(* IEC 61131-3 sources: volt/packages/volt-lsp-iec/test-corpus/lenze-mid/Device/Plc Logic/Application/Library Manager/L_TT1P_TechnologyModules (part 4) *)

(* ---- L_MB1P_POSPROFILER.pou ---- *)
FUNCTION_BLOCK L_MB1P_POSPROFILER
VAR_INPUT
	XEXECUTE : BOOL;
	XAUXEXECUTE : BOOL;
	XABORT : BOOL;
	XPOSMODE : BOOL;
	ROVERRIDESPEED : REAL;
	ROVERRIDEACC : REAL;
	ROVERRIDEDEC : REAL;
	ROVERRIDEJERKACC : REAL;
	ROVERRIDEJERKDEC : REAL;
	LRACTPOS : LREAL;
	LRACTSPEED : LREAL;
	LRACTACC : LREAL;
	RTASKCYCLE : REAL;
END_VAR
VAR_OUTPUT
	XBUSY : BOOL;
	XDONE : BOOL;
	XABORTED : BOOL;
	XERROR : BOOL;
	LRSETPOS : LREAL;
	LRSETSPEED : LREAL;
	LRSETACC : LREAL;
	DWSTATE : DWORD;
	DWPROFILETYPE : DWORD;
END_VAR
VAR_IN_OUT
	SCPROFILEPARAMETER : L_MB1P_ProfileParameter;
END_VAR
VAR
	SCPROFILEDATA : L_MB1P_ProfileData;
	LREVALTIME : LREAL;
	DWSTATEOFINTERPOLATOR : DWORD;
	XFLAGEXECUTE : BOOL;
	XFLAGAUXEXECUTE : BOOL;
	XFLAGABORT : BOOL;
	SCPROFILEPARAMETERINT : L_MB1P_ProfileParameter;
	ROVERRIDESPEEDOLD : REAL;
	ROVERRIDEACCOLD : REAL;
	ROVERRIDEDECOLD : REAL;
	ROVERRIDEJERKACCOLD : REAL;
	ROVERRIDEJERKDECOLD : REAL;
	XSTARTCALCPROF : BOOL;
	XVELOVEREQZERO : BOOL;
	ARG1 : LREAL;
END_VAR
END_FUNCTION_BLOCK

METHOD CALCPROFILE : BOOL
VAR_INPUT
	DWPROFILETYPE : DWORD;
	LRSTARTACC : LREAL;
	LRSTARTVEL : LREAL;
	SCPROFILEPARAMETER : L_MB1P_ProfileParameter;
	SCMINPROFILEDATA : L_MB1P_IntProfileData;
	SCMAXPROFILEDATA : L_MB1P_IntProfileData;
END_VAR
VAR_OUTPUT
	SCPROFILEDATA : L_MB1P_ProfileData;
	DWSTATE : DWORD;
END_VAR
END_METHOD

METHOD CALCPROFILEDATA : BOOL
VAR_INPUT
	LRSTARTACC : LREAL;
	LRSTARTVEL : LREAL;
	LRSTARTPOS : LREAL;
	XVELMODE : BOOL;
END_VAR
VAR_OUTPUT
	XERROR : BOOL;
	DWSTATE : DWORD;
	DWPROFILETYPE : DWORD;
END_VAR
VAR_IN_OUT
	SCPROFILEDATA : L_MB1P_ProfileData;
	SCPROFILEPARAMETER : L_MB1P_ProfileParameter;
END_VAR
END_METHOD

METHOD IDENTPROFILETYPE : DWORD
VAR_INPUT
	XVELMODE : BOOL;
	LRSTARTACC : LREAL;
	LRSTARTVEL : LREAL;
	SCPROFILEPARAMETER : L_MB1P_ProfileParameter;
END_VAR
VAR_OUTPUT
	DWPROFILETYPE : DWORD;
	SCMINPROFILEDATA : L_MB1P_IntProfileData;
	SCMAXPROFILEDATA : L_MB1P_IntProfileData;
	DWSTATE : DWORD;
END_VAR
END_METHOD

METHOD PROFILEINTERPOLATOR : BOOL
VAR_INPUT
	LREVALTIME : LREAL;
END_VAR
VAR_OUTPUT
	DWSTATE : DWORD;
	LRSETPOS : LREAL;
	LRSETVEL : LREAL;
	LRSETACC : LREAL;
END_VAR
VAR_IN_OUT
	SCPROFILEDATA : L_MB1P_ProfileData;
END_VAR
END_METHOD

METHOD RESETOUTPUT
END_METHOD

METHOD CALCSQRT : LREAL
VAR_INPUT
	ARG1 : LREAL;
END_VAR
END_METHOD

METHOD CALCMINPOSPROFILE : BOOL
VAR_INPUT
	MAXVEL : LREAL;
	MAXACC1 : LREAL;
	MAXACC2 : LREAL;
	JERKACC1 : LREAL;
	JERKACC2 : LREAL;
	RECIPRJERKACC1 : LREAL;
	RECIPRJERKACC2 : LREAL;
	V0_ACC1 : LREAL;
	V0_ACC2 : LREAL;
	A0_ACC1 : LREAL;
	A0_ACC2 : LREAL;
END_VAR
VAR_OUTPUT
	DIMINPOSPROFILETYPE : DINT;
	MINPOSPROFILEDATA : L_MB1P_IntProfileData;
	VMAXMINTRIACC1 : LREAL;
	VMAX_MINTRIACC2 : LREAL;
END_VAR
END_METHOD

METHOD CALCMINPROFILENEGACC : BOOL
VAR_INPUT
	VMAX : LREAL;
	AMAX : LREAL;
	V0 : LREAL;
	A0 : LREAL;
	JERK : LREAL;
	JERKRECIPR : LREAL;
END_VAR
VAR_OUTPUT
	DWPROFILETYPE : DWORD;
	PROFILEDATA_NEGACC : L_MB1P_IntProfileDataAcc;
END_VAR
END_METHOD

METHOD CALCMINPROFILEPOSACC : BOOL
VAR_INPUT
	VMAX : LREAL;
	AMAX : LREAL;
	V0 : LREAL;
	A0 : LREAL;
	JERK : LREAL;
	JERKRECIPR : LREAL;
END_VAR
VAR_OUTPUT
	DWPROFILETYPE : DWORD;
	PROFILEDATA_POSACC : L_MB1P_IntProfileDataAcc;
END_VAR
END_METHOD

METHOD CALCMINTRI : BOOL
VAR_INPUT
	RECIPRJERKACC1 : LREAL;
	RECIPRJERKACC2 : LREAL;
	A0_ACC1 : LREAL;
	V0_ACC1 : LREAL;
	A0_ACC2 : LREAL;
	V0_ACC2 : LREAL;
END_VAR
VAR_OUTPUT
	VMAXMINTRIACC1 : LREAL;
	VMAXMINTRIACC2 : LREAL;
	PROFILEDATA_ACC1 : L_MB1P_IntProfileDataAcc;
	PROFILEDATA_ACC2 : L_MB1P_IntProfileDataAcc;
END_VAR
END_METHOD

METHOD CHECKPROFILEDATA
VAR_INPUT
	DWMODE : DWORD;
	LRTARGETPOS : LREAL;
	LRTARGETVEL : LREAL;
	LRTARGETACC : LREAL;
	LRJERKPHASE7 : LREAL;
END_VAR
VAR_OUTPUT
	XERROR : BOOL;
END_VAR
VAR_IN_OUT
	SCPROFILEDATA : L_MB1P_ProfileData;
END_VAR
END_METHOD

METHOD IDENTMINNEGPROFILE : BOOL
VAR_INPUT
	MINPOSPROFILETYPE : DINT;
	MAXVEL : LREAL;
	MAXACC : LREAL;
	JERK : LREAL;
	RECIPRJERK : LREAL;
	V0_ACC1 : LREAL;
	V0_ACC2 : LREAL;
	A0_ACC1 : LREAL;
	A0_ACC2 : LREAL;
	TARGETPOS : LREAL;
END_VAR
VAR_OUTPUT
	DWPROFILETYPE : DWORD;
END_VAR
VAR_IN_OUT
	SCMAXPROFILEDATA : L_MB1P_IntProfileData;
	SCMINPROFILEDATA : L_MB1P_IntProfileData;
END_VAR
END_METHOD

METHOD IDENTMINPOSPROFILE : BOOL
VAR_INPUT
	MAXVEL : LREAL;
	MAXACC1 : LREAL;
	MAXACC2 : LREAL;
	JERKACC1 : LREAL;
	JERKACC2 : LREAL;
	V0_ACC1 : LREAL;
	V0_ACC2 : LREAL;
	A0_ACC1 : LREAL;
	A0_ACC2 : LREAL;
	TARGETPOS : LREAL;
END_VAR
VAR_OUTPUT
	DWPROFILETYPE : DWORD;
	SCMAXPROFILEDATA : L_MB1P_IntProfileData;
	SCMINPROFILEDATA : L_MB1P_IntProfileData;
END_VAR
END_METHOD

METHOD IDENTSIMPLETRAPNEG : BOOL
VAR_INPUT
	MAXACC2 : LREAL;
	V0_ACC1 : LREAL;
	V0_ACC2 : LREAL;
	A0_ACC1 : LREAL;
	A0_ACC2 : LREAL;
	JERKACC1 : LREAL;
	JERKACC2 : LREAL;
	RECIPRJERKACC2 : LREAL;
	TARGETPOS : LREAL;
END_VAR
VAR_OUTPUT
	DWPROFILETYPE : DWORD;
END_VAR
VAR_IN_OUT
	SCMINPROFILEDATA : L_MB1P_IntProfileData;
	SCMAXPROFILEDATA : L_MB1P_IntProfileData;
END_VAR
END_METHOD

METHOD IDENTSIMPLETRAPPOSTRINEG : BOOL
VAR_INPUT
	MAXACC1 : LREAL;
	JERKACC1 : LREAL;
	RECIPRJERKACC1 : LREAL;
	V0_ACC1 : LREAL;
	A0_ACC1 : LREAL;
	VMAXMINTRIACC1 : LREAL;
	VMAXMINTRIACC2 : LREAL;
	JERKACC2 : LREAL;
	TARGETPOS : LREAL;
END_VAR
VAR_OUTPUT
	DWPROFILETYPE : DWORD;
END_VAR
VAR_IN_OUT
	SCMINPROFILEDATA : L_MB1P_IntProfileData;
	SCMAXPROFILEDATA : L_MB1P_IntProfileData;
END_VAR
END_METHOD

METHOD IDENTSIMPLETRINEG : BOOL
VAR_INPUT
	V0_ACC1 : LREAL;
	A0_ACC1 : LREAL;
	A0_ACC2 : LREAL;
	JERKACC1 : LREAL;
	JERKACC2 : LREAL;
	RECIPRJERKACC2 : LREAL;
	TARGETPOS : LREAL;
END_VAR
VAR_OUTPUT
	DWPROFILETYPE : DWORD;
END_VAR
VAR_IN_OUT
	SCMINPROFILEDATA : L_MB1P_IntProfileData;
	SCMAXPROFILEDATA : L_MB1P_IntProfileData;
END_VAR
END_METHOD

METHOD IDENTSIMPLETRIPOSTRAPNEG : BOOL
VAR_INPUT
	MAXACC2 : LREAL;
	JERKACC2 : LREAL;
	RECIPRJERKACC2 : LREAL;
	V0_ACC2 : LREAL;
	A0_ACC2 : LREAL;
	VMAXMINTRIACC1 : LREAL;
	JERKACC1 : LREAL;
	TARGETPOS : LREAL;
END_VAR
VAR_OUTPUT
	DWPROFILETYPE : DWORD;
END_VAR
VAR_IN_OUT
	SCMINPROFILEDATA : L_MB1P_IntProfileData;
	SCMAXPROFILEDATA : L_MB1P_IntProfileData;
END_VAR
END_METHOD

METHOD IDENTSIMPLETRIPOSTRINEG : BOOL
VAR_INPUT
	V0_ACC1 : LREAL;
	A0_ACC1 : LREAL;
	AMAX : LREAL;
	RECIPRJERKACC1 : LREAL;
	JERKACC1 : LREAL;
	JERKACC2 : LREAL;
	TARGETPOS : LREAL;
	VMAXMINTRIACC1 : LREAL;
	VMAXMINTRIACC2 : LREAL;
END_VAR
VAR_OUTPUT
	DWPROFILETYPE : DWORD;
END_VAR
VAR_IN_OUT
	SCMINPROFILEDATA : L_MB1P_IntProfileData;
	SCMAXPROFILEDATA : L_MB1P_IntProfileData;
END_VAR
END_METHOD

METHOD IDENTTRAPTRI : BOOL
VAR_INPUT
	V_MINTRAPEZACC1 : LREAL;
	MAXACC1 : LREAL;
	JERKACC1 : LREAL;
	JERKACC2 : LREAL;
	A0_ACC1 : LREAL;
	A0_ACC2 : LREAL;
	V0_ACC1 : LREAL;
	V0_ACC2 : LREAL;
	T1_ACC1 : LREAL;
	T3_ACC1 : LREAL;
	DS_1_ACC1 : LREAL;
	TARGETPOS : LREAL;
END_VAR
VAR_OUTPUT
	DWPROFILETYPE : DWORD;
END_VAR
VAR_IN_OUT
	SCMINPROFILEDATA : L_MB1P_IntProfileData;
	SCMAXPROFILEDATA : L_MB1P_IntProfileData;
END_VAR
END_METHOD

METHOD IDENTTRITRAP : BOOL
VAR_INPUT
	V_MINTRAPEZACC2 : LREAL;
	MAXACC2 : LREAL;
	JERKACC1 : LREAL;
	JERKACC2 : LREAL;
	A0_ACC1 : LREAL;
	A0_ACC2 : LREAL;
	V0_ACC1 : LREAL;
	V0_ACC2 : LREAL;
	T1_ACC2 : LREAL;
	T3_ACC2 : LREAL;
	DS_1_ACC2 : LREAL;
	TARGETPOS : LREAL;
END_VAR
VAR_OUTPUT
	DWPROFILETYPE : DWORD;
END_VAR
VAR_IN_OUT
	SCMINPROFILEDATA : L_MB1P_IntProfileData;
	SCMAXPROFILEDATA : L_MB1P_IntProfileData;
END_VAR
END_METHOD

METHOD CALCPROFILE_10A0 : BOOL
VAR_INPUT
	LRSTARTACC : LREAL;
	LRSTARTVEL : LREAL;
	LRMAXACC : LREAL;
	LRMAXDEC : LREAL;
	LRMAXVEL : LREAL;
	LRTARGETACC : LREAL;
	LRTARGETVEL : LREAL;
	LRTARGETPOS : LREAL;
	LRJERKACC : LREAL;
	LRJERKDEC : LREAL;
	LRJERKTIMEACC : LREAL;
	LRJERKTIMEDEC : LREAL;
END_VAR
VAR_OUTPUT
	DWSTATE : DWORD;
END_VAR
VAR_IN_OUT
	SCPROFILEDATA : L_MB1P_ProfileData;
	SCPROFILEPARAMETER : L_MB1P_ProfileParameter;
END_VAR
END_METHOD

METHOD CALCPROFILE_10A0_A0GTAMAX : BOOL
VAR_INPUT
	LRSTARTACC : LREAL;
	LRSTARTVEL : LREAL;
	LRMAXACC : LREAL;
	LRMAXVEL : LREAL;
	LRMAXDEC : LREAL;
	LRTARGETACC : LREAL;
	LRTARGETVEL : LREAL;
	LRTARGETPOS : LREAL;
	LRJERKTIMEACC : LREAL;
	LRJERKTIMEDEC : LREAL;
	LRJERKACC : LREAL;
	LRJERKDEC : LREAL;
END_VAR
VAR_IN_OUT
	SCPROFILEDATA : L_MB1P_ProfileData;
END_VAR
END_METHOD

METHOD CALCPROFILE_10A0_A0LTAMAX : BOOL
VAR_INPUT
	LRSTARTACC : LREAL;
	LRSTARTVEL : LREAL;
	LRMAXACC : LREAL;
	LRMAXVEL : LREAL;
	LRMAXDEC : LREAL;
	LRTARGETACC : LREAL;
	LRTARGETVEL : LREAL;
	LRTARGETPOS : LREAL;
	LRJERKTIMEACC : LREAL;
	LRJERKTIMEDEC : LREAL;
	LRJERKACC : LREAL;
	LRJERKDEC : LREAL;
END_VAR
VAR_IN_OUT
	SCPROFILEDATA : L_MB1P_ProfileData;
END_VAR
END_METHOD

METHOD CALCPROFILE_10B0 : BOOL
VAR_INPUT
	LRSTARTACC : LREAL;
	LRSTARTVEL : LREAL;
	LRMAXACC : LREAL;
	LRMAXDEC : LREAL;
	LRMAXVEL : LREAL;
	LRTARGETACC : LREAL;
	LRTARGETVEL : LREAL;
	LRTARGETPOS : LREAL;
	LRJERKACC : LREAL;
	LRJERKDEC : LREAL;
	LRJERKTIMEACC : LREAL;
	LRJERKTIMEDEC : LREAL;
END_VAR
VAR_OUTPUT
	DWSTATE : DWORD;
END_VAR
VAR_IN_OUT
	SCPROFILEDATA : L_MB1P_ProfileData;
	SCPROFILEPARAMETER : L_MB1P_ProfileParameter;
END_VAR
END_METHOD

METHOD CALCPROFILE_10B0_A0GTAMAX : BOOL
VAR_INPUT
	LRSTARTACC : LREAL;
	LRSTARTVEL : LREAL;
	LRMAXACC : LREAL;
	LRMAXVEL : LREAL;
	LRMAXDEC : LREAL;
	LRTARGETACC : LREAL;
	LRTARGETVEL : LREAL;
	LRTARGETPOS : LREAL;
	LRJERKTIMEACC : LREAL;
	LRJERKTIMEDEC : LREAL;
	LRJERKACC : LREAL;
	LRJERKDEC : LREAL;
END_VAR
VAR_IN_OUT
	SCPROFILEDATA : L_MB1P_ProfileData;
END_VAR
END_METHOD

METHOD CALCPROFILE_10B0_A0LTAMAX : BOOL
VAR_INPUT
	LRSTARTACC : LREAL;
	LRSTARTVEL : LREAL;
	LRMAXACC : LREAL;
	LRMAXVEL : LREAL;
	LRMAXDEC : LREAL;
	LRTARGETACC : LREAL;
	LRTARGETVEL : LREAL;
	LRTARGETPOS : LREAL;
	LRJERKTIMEACC : LREAL;
	LRJERKTIMEDEC : LREAL;
	LRJERKACC : LREAL;
	LRJERKDEC : LREAL;
END_VAR
VAR_IN_OUT
	SCPROFILEDATA : L_MB1P_ProfileData;
END_VAR
END_METHOD

METHOD CALCPROFILE_10C0 : BOOL
VAR_INPUT
	LRSTARTACC : LREAL;
	LRSTARTVEL : LREAL;
	LRMAXACC : LREAL;
	LRMAXDEC : LREAL;
	LRMAXVEL : LREAL;
	LRTARGETACC : LREAL;
	LRTARGETVEL : LREAL;
	LRTARGETPOS : LREAL;
	LRJERKACC : LREAL;
	LRJERKDEC : LREAL;
	LRJERKTIMEACC : LREAL;
	LRJERKTIMEDEC : LREAL;
END_VAR
VAR_OUTPUT
	DWSTATE : DWORD;
END_VAR
VAR_IN_OUT
	SCPROFILEDATA : L_MB1P_ProfileData;
	SCPROFILEPARAMETER : L_MB1P_ProfileParameter;
END_VAR
END_METHOD

METHOD CALCPROFILE_10C0_A0LTAMAXT31 : BOOL
VAR_INPUT
	LRSTARTACC : LREAL;
	LRSTARTVEL : LREAL;
	LRMAXACC : LREAL;
	LRMAXVEL : LREAL;
	LRMAXDEC : LREAL;
	LRTARGETACC : LREAL;
	LRTARGETVEL : LREAL;
	LRTARGETPOS : LREAL;
	LRJERKTIMEACC : LREAL;
	LRJERKTIMEDEC : LREAL;
	LRJERKACC : LREAL;
	LRJERKDEC : LREAL;
END_VAR
VAR_IN_OUT
	SCPROFILEDATA : L_MB1P_ProfileData;
END_VAR
END_METHOD

METHOD CALCPROFILE_10C0_A0LTAMAXT32 : BOOL
VAR_INPUT
	LRSTARTACC : LREAL;
	LRSTARTVEL : LREAL;
	LRMAXACC : LREAL;
	LRMAXVEL : LREAL;
	LRMAXDEC : LREAL;
	LRTARGETACC : LREAL;
	LRTARGETVEL : LREAL;
	LRTARGETPOS : LREAL;
	LRJERKTIMEACC : LREAL;
	LRJERKTIMEDEC : LREAL;
	LRJERKACC : LREAL;
	LRJERKDEC : LREAL;
END_VAR
VAR_IN_OUT
	SCPROFILEDATA : L_MB1P_ProfileData;
END_VAR
END_METHOD

METHOD CALCPROFILE_10D0 : BOOL
VAR_INPUT
	LRSTARTACC : LREAL;
	LRSTARTVEL : LREAL;
	LRMAXACC : LREAL;
	LRMAXDEC : LREAL;
	LRMAXVEL : LREAL;
	LRTARGETACC : LREAL;
	LRTARGETVEL : LREAL;
	LRTARGETPOS : LREAL;
	LRJERKACC : LREAL;
	LRJERKDEC : LREAL;
	LRJERKTIMEACC : LREAL;
	LRJERKTIMEDEC : LREAL;
END_VAR
VAR_OUTPUT
	DWSTATE : DWORD;
END_VAR
VAR_IN_OUT
	SCPROFILEDATA : L_MB1P_ProfileData;
	SCPROFILEPARAMETER : L_MB1P_ProfileParameter;
END_VAR
END_METHOD

METHOD CALCPROFILE_10D0_A0LTAMAXT31T51 : BOOL
VAR_INPUT
	LRSTARTACC : LREAL;
	LRSTARTVEL : LREAL;
	LRMAXACC : LREAL;
	LRMAXVEL : LREAL;
	LRMAXDEC : LREAL;
	LRTARGETACC : LREAL;
	LRTARGETVEL : LREAL;
	LRTARGETPOS : LREAL;
	LRJERKTIMEACC : LREAL;
	LRJERKTIMEDEC : LREAL;
	LRJERKACC : LREAL;
	LRJERKDEC : LREAL;
END_VAR
VAR_IN_OUT
	SCPROFILEDATA : L_MB1P_ProfileData;
END_VAR
END_METHOD

METHOD CALCPROFILE_10D0_A0LTAMAXT31T52 : BOOL
VAR_INPUT
	LRSTARTACC : LREAL;
	LRSTARTVEL : LREAL;
	LRMAXACC : LREAL;
	LRMAXVEL : LREAL;
	LRMAXDEC : LREAL;
	LRTARGETACC : LREAL;
	LRTARGETVEL : LREAL;
	LRTARGETPOS : LREAL;
	LRJERKTIMEACC : LREAL;
	LRJERKTIMEDEC : LREAL;
	LRJERKACC : LREAL;
	LRJERKDEC : LREAL;
END_VAR
VAR_IN_OUT
	SCPROFILEDATA : L_MB1P_ProfileData;
END_VAR
END_METHOD

METHOD CALCPROFILE_10D0_A0LTAMAXT32T51 : BOOL
VAR_INPUT
	LRSTARTACC : LREAL;
	LRSTARTVEL : LREAL;
	LRMAXACC : LREAL;
	LRMAXVEL : LREAL;
	LRMAXDEC : LREAL;
	LRTARGETACC : LREAL;
	LRTARGETVEL : LREAL;
	LRTARGETPOS : LREAL;
	LRJERKTIMEACC : LREAL;
	LRJERKTIMEDEC : LREAL;
	LRJERKACC : LREAL;
	LRJERKDEC : LREAL;
END_VAR
VAR_IN_OUT
	SCPROFILEDATA : L_MB1P_ProfileData;
END_VAR
END_METHOD

METHOD CALCPROFILE_10D0_A0LTAMAXT32T52 : BOOL
VAR_INPUT
	LRSTARTACC : LREAL;
	LRSTARTVEL : LREAL;
	LRMAXACC : LREAL;
	LRMAXVEL : LREAL;
	LRMAXDEC : LREAL;
	LRTARGETACC : LREAL;
	LRTARGETVEL : LREAL;
	LRTARGETPOS : LREAL;
	LRJERKTIMEACC : LREAL;
	LRJERKTIMEDEC : LREAL;
	LRJERKACC : LREAL;
	LRJERKDEC : LREAL;
END_VAR
VAR_IN_OUT
	SCPROFILEDATA : L_MB1P_ProfileData;
END_VAR
END_METHOD

METHOD CALCPROFILE_20A0 : BOOL
VAR_INPUT
	LRSTARTACC : LREAL;
	LRSTARTVEL : LREAL;
	LRMAXACC : LREAL;
	LRMAXDEC : LREAL;
	LRMAXVEL : LREAL;
	LRTARGETACC : LREAL;
	LRTARGETVEL : LREAL;
	LRTARGETPOS : LREAL;
	LRJERKACC : LREAL;
	LRJERKDEC : LREAL;
	LRJERKTIMEACC : LREAL;
	LRJERKTIMEDEC : LREAL;
END_VAR
VAR_OUTPUT
	DWSTATE : DWORD;
END_VAR
VAR_IN_OUT
	SCPROFILEDATA : L_MB1P_ProfileData;
	SCPROFILEPARAMETER : L_MB1P_ProfileParameter;
END_VAR
END_METHOD

METHOD CALCPROFILE_20A0_A0GTAMAXT71 : BOOL
VAR_INPUT
	LRSTARTACC : LREAL;
	LRSTARTVEL : LREAL;
	LRMAXACC : LREAL;
	LRMAXDEC : LREAL;
	LRMAXVEL : LREAL;
	LRTARGETACC : LREAL;
	LRTARGETVEL : LREAL;
	LRTARGETPOS : LREAL;
	LRJERKACC : LREAL;
	LRJERKDEC : LREAL;
	LRJERKTIMEACC : LREAL;
	LRJERKTIMEDEC : LREAL;
END_VAR
VAR_IN_OUT
	SCPROFILEDATA : L_MB1P_ProfileData;
END_VAR
END_METHOD

METHOD CALCPROFILE_20A0_A0GTAMAXT72 : BOOL
VAR_INPUT
	LRSTARTACC : LREAL;
	LRSTARTVEL : LREAL;
	LRMAXACC : LREAL;
	LRMAXDEC : LREAL;
	LRMAXVEL : LREAL;
	LRTARGETACC : LREAL;
	LRTARGETVEL : LREAL;
	LRTARGETPOS : LREAL;
	LRJERKACC : LREAL;
	LRJERKDEC : LREAL;
	LRJERKTIMEACC : LREAL;
	LRJERKTIMEDEC : LREAL;
END_VAR
VAR_IN_OUT
	SCPROFILEDATA : L_MB1P_ProfileData;
END_VAR
END_METHOD

METHOD CALCPROFILE_20A0_A0LTAMAXT71 : BOOL
VAR_INPUT
	LRSTARTACC : LREAL;
	LRSTARTVEL : LREAL;
	LRMAXACC : LREAL;
	LRMAXDEC : LREAL;
	LRMAXVEL : LREAL;
	LRTARGETACC : LREAL;
	LRTARGETVEL : LREAL;
	LRTARGETPOS : LREAL;
	LRJERKACC : LREAL;
	LRJERKDEC : LREAL;
	LRJERKTIMEACC : LREAL;
	LRJERKTIMEDEC : LREAL;
END_VAR
VAR_IN_OUT
	SCPROFILEDATA : L_MB1P_ProfileData;
END_VAR
END_METHOD

METHOD CALCPROFILE_20A0_A0LTAMAXT72 : BOOL
VAR_INPUT
	LRSTARTACC : LREAL;
	LRSTARTVEL : LREAL;
	LRMAXACC : LREAL;
	LRMAXDEC : LREAL;
	LRMAXVEL : LREAL;
	LRTARGETACC : LREAL;
	LRTARGETVEL : LREAL;
	LRTARGETPOS : LREAL;
	LRJERKACC : LREAL;
	LRJERKDEC : LREAL;
	LRJERKTIMEACC : LREAL;
	LRJERKTIMEDEC : LREAL;
END_VAR
VAR_IN_OUT
	SCPROFILEDATA : L_MB1P_ProfileData;
END_VAR
END_METHOD

METHOD CALCPROFILE_20B0 : BOOL
VAR_INPUT
	LRSTARTACC : LREAL;
	LRSTARTVEL : LREAL;
	LRMAXACC : LREAL;
	LRMAXDEC : LREAL;
	LRMAXVEL : LREAL;
	LRTARGETACC : LREAL;
	LRTARGETVEL : LREAL;
	LRTARGETPOS : LREAL;
	LRJERKACC : LREAL;
	LRJERKDEC : LREAL;
	LRJERKTIMEACC : LREAL;
	LRJERKTIMEDEC : LREAL;
	SCMAXPROFILEDATA : L_MB1P_IntProfileData;
	SCMINPROFILEDATA : L_MB1P_IntProfileData;
END_VAR
VAR_OUTPUT
	DWSTATE : DWORD;
END_VAR
VAR_IN_OUT
	SCPROFILEDATA : L_MB1P_ProfileData;
	SCPROFILEPARAMETER : L_MB1P_ProfileParameter;
END_VAR
END_METHOD

METHOD CALCPROFILE_20B0_A0GTAMAXSEARCHTIMEST5T7 : BOOL
VAR_INPUT
	LRSTARTACC : LREAL;
	LRSTARTVEL : LREAL;
	LRMAXACC : LREAL;
	LRMAXDEC : LREAL;
	LRMAXVEL : LREAL;
	LRTARGETACC : LREAL;
	LRTARGETVEL : LREAL;
	LRTARGETPOS : LREAL;
	LRJERKACC : LREAL;
	LRJERKDEC : LREAL;
	LRJERKTIMEACC : LREAL;
	LRJERKTIMEDEC : LREAL;
	T5_STARTVALUE : LREAL;
	T7_STARTVALUE : LREAL;
END_VAR
VAR_OUTPUT
	T5 : LREAL;
	T7 : LREAL;
END_VAR
END_METHOD

METHOD CALCPROFILE_20B0_A0GTAMAXT5T7 : BOOL
VAR_INPUT
	LRSTARTACC : LREAL;
	LRSTARTVEL : LREAL;
	LRMAXACC : LREAL;
	LRMAXDEC : LREAL;
	LRMAXVEL : LREAL;
	LRTARGETACC : LREAL;
	LRTARGETVEL : LREAL;
	LRTARGETPOS : LREAL;
	LRJERKACC : LREAL;
	LRJERKDEC : LREAL;
	LRJERKTIMEACC : LREAL;
	LRJERKTIMEDEC : LREAL;
	T5 : LREAL;
	T7 : LREAL;
END_VAR
VAR_IN_OUT
	SCPROFILEDATA : L_MB1P_ProfileData;
END_VAR
END_METHOD

METHOD CALCPROFILE_20B0_A0LTAMAXSEARCHTIMEST5T7 : BOOL
VAR_INPUT
	LRSTARTACC : LREAL;
	LRSTARTVEL : LREAL;
	LRMAXACC : LREAL;
	LRMAXDEC : LREAL;
	LRMAXVEL : LREAL;
	LRTARGETACC : LREAL;
	LRTARGETVEL : LREAL;
	LRTARGETPOS : LREAL;
	LRJERKACC : LREAL;
	LRJERKDEC : LREAL;
	LRJERKTIMEACC : LREAL;
	LRJERKTIMEDEC : LREAL;
	T5_STARTVALUE : LREAL;
	T7_STARTVALUE : LREAL;
END_VAR
VAR_OUTPUT
	T5 : LREAL;
	T7 : LREAL;
END_VAR
END_METHOD

METHOD CALCPROFILE_20B0_A0LTAMAXT5T7 : BOOL
VAR_INPUT
	LRSTARTACC : LREAL;
	LRSTARTVEL : LREAL;
	LRMAXACC : LREAL;
	LRMAXDEC : LREAL;
	LRMAXVEL : LREAL;
	LRTARGETACC : LREAL;
	LRTARGETVEL : LREAL;
	LRTARGETPOS : LREAL;
	LRJERKACC : LREAL;
	LRJERKDEC : LREAL;
	LRJERKTIMEACC : LREAL;
	LRJERKTIMEDEC : LREAL;
	T5 : LREAL;
	T7 : LREAL;
END_VAR
VAR_IN_OUT
	SCPROFILEDATA : L_MB1P_ProfileData;
END_VAR
END_METHOD

METHOD CALCPROFILE_20BA : BOOL
VAR_INPUT
	LRSTARTACC : LREAL;
	LRSTARTVEL : LREAL;
	LRMAXACC : LREAL;
	LRMAXDEC : LREAL;
	LRMAXVEL : LREAL;
	LRTARGETACC : LREAL;
	LRTARGETVEL : LREAL;
	LRTARGETPOS : LREAL;
	LRJERKACC : LREAL;
	LRJERKDEC : LREAL;
	LRJERKTIMEACC : LREAL;
	LRJERKTIMEDEC : LREAL;
	SCMAXPROFILEDATA : L_MB1P_IntProfileData;
	SCMINPROFILEDATA : L_MB1P_IntProfileData;
END_VAR
VAR_OUTPUT
	DWSTATE : DWORD;
END_VAR
VAR_IN_OUT
	SCPROFILEDATA : L_MB1P_ProfileData;
	SCPROFILEPARAMETER : L_MB1P_ProfileParameter;
END_VAR
END_METHOD

METHOD CALCPROFILE_20BA_A0GTAMAX : BOOL
VAR_INPUT
	LRSTARTACC : LREAL;
	LRSTARTVEL : LREAL;
	LRMAXACC : LREAL;
	LRMAXDEC : LREAL;
	LRMAXVEL : LREAL;
	LRTARGETACC : LREAL;
	LRTARGETVEL : LREAL;
	LRTARGETPOS : LREAL;
	LRJERKACC : LREAL;
	LRJERKDEC : LREAL;
	LRJERKTIMEACC : LREAL;
	LRJERKTIMEDEC : LREAL;
	T7 : LREAL;
END_VAR
VAR_IN_OUT
	SCPROFILEDATA : L_MB1P_ProfileData;
END_VAR
END_METHOD

METHOD CALCPROFILE_20BA_A0LETAMAX : BOOL
VAR_INPUT
	LRSTARTACC : LREAL;
	LRSTARTVEL : LREAL;
	LRMAXACC : LREAL;
	LRMAXDEC : LREAL;
	LRMAXVEL : LREAL;
	LRTARGETACC : LREAL;
	LRTARGETVEL : LREAL;
	LRTARGETPOS : LREAL;
	LRJERKACC : LREAL;
	LRJERKDEC : LREAL;
	LRJERKTIMEACC : LREAL;
	LRJERKTIMEDEC : LREAL;
	T7 : LREAL;
END_VAR
VAR_IN_OUT
	SCPROFILEDATA : L_MB1P_ProfileData;
END_VAR
END_METHOD

METHOD CALCPROFILE_20BA_AOGTAMAX_SEARCHTIMES : BOOL
VAR_INPUT
	LRSTARTACC : LREAL;
	LRSTARTVEL : LREAL;
	LRMAXACC : LREAL;
	LRMAXDEC : LREAL;
	LRMAXVEL : LREAL;
	LRTARGETACC : LREAL;
	LRTARGETVEL : LREAL;
	LRTARGETPOS : LREAL;
	LRJERKACC : LREAL;
	LRJERKDEC : LREAL;
	LRJERKTIMEACC : LREAL;
	LRJERKTIMEDEC : LREAL;
	T7_MINVALUE : LREAL;
	T7_MAXVALUE : LREAL;
END_VAR
VAR_OUTPUT
	T7 : LREAL;
END_VAR
END_METHOD

METHOD CALCPROFILE_20BA_AOLETAMAX_SEARCHTIMES : BOOL
VAR_INPUT
	LRSTARTACC : LREAL;
	LRSTARTVEL : LREAL;
	LRMAXACC : LREAL;
	LRMAXDEC : LREAL;
	LRMAXVEL : LREAL;
	LRTARGETACC : LREAL;
	LRTARGETVEL : LREAL;
	LRTARGETPOS : LREAL;
	LRJERKACC : LREAL;
	LRJERKDEC : LREAL;
	LRJERKTIMEACC : LREAL;
	LRJERKTIMEDEC : LREAL;
	T7_MINVALUE : LREAL;
	T7_MAXVALUE : LREAL;
END_VAR
VAR_OUTPUT
	T7 : LREAL;
END_VAR
END_METHOD

METHOD CALCPROFILE_20C0 : BOOL
VAR_INPUT
	LRSTARTACC : LREAL;
	LRSTARTVEL : LREAL;
	LRMAXACC : LREAL;
	LRMAXDEC : LREAL;
	LRMAXVEL : LREAL;
	LRTARGETACC : LREAL;
	LRTARGETVEL : LREAL;
	LRTARGETPOS : LREAL;
	LRJERKACC : LREAL;
	LRJERKDEC : LREAL;
	LRJERKTIMEACC : LREAL;
	LRJERKTIMEDEC : LREAL;
	SCMAXPROFILEDATA : L_MB1P_IntProfileData;
	SCMINPROFILEDATA : L_MB1P_IntProfileData;
END_VAR
VAR_OUTPUT
	DWSTATE : DWORD;
END_VAR
VAR_IN_OUT
	SCPROFILEDATA : L_MB1P_ProfileData;
	SCPROFILEPARAMETER : L_MB1P_ProfileParameter;
END_VAR
END_METHOD

METHOD CALCPROFILE_20C0_SEARCHTIMEST5T7 : BOOL
VAR_INPUT
	LRSTARTACC : LREAL;
	LRSTARTVEL : LREAL;
	LRMAXACC : LREAL;
	LRMAXDEC : LREAL;
	LRMAXVEL : LREAL;
	LRTARGETACC : LREAL;
	LRTARGETVEL : LREAL;
	LRTARGETPOS : LREAL;
	LRJERKACC : LREAL;
	LRJERKDEC : LREAL;
	LRJERKTIMEACC : LREAL;
	LRJERKTIMEDEC : LREAL;
	T5_STARTVALUE : LREAL;
	T7_STARTVALUE : LREAL;
END_VAR
VAR_OUTPUT
	T5 : LREAL;
	T7 : LREAL;
END_VAR
END_METHOD

METHOD CALCPROFILE_20C0_AELTAMAXT5T7 : BOOL
VAR_INPUT
	LRSTARTACC : LREAL;
	LRSTARTVEL : LREAL;
	LRMAXACC : LREAL;
	LRMAXDEC : LREAL;
	LRMAXVEL : LREAL;
	LRTARGETACC : LREAL;
	LRTARGETVEL : LREAL;
	LRTARGETPOS : LREAL;
	LRJERKACC : LREAL;
	LRJERKDEC : LREAL;
	LRJERKTIMEACC : LREAL;
	LRJERKTIMEDEC : LREAL;
	T5 : LREAL;
	T7 : LREAL;
END_VAR
VAR_IN_OUT
	SCPROFILEDATA : L_MB1P_ProfileData;
END_VAR
END_METHOD

METHOD CALCPROFILE_20CB : BOOL
VAR_INPUT
	LRSTARTACC : LREAL;
	LRSTARTVEL : LREAL;
	LRMAXACC : LREAL;
	LRMAXDEC : LREAL;
	LRMAXVEL : LREAL;
	LRTARGETACC : LREAL;
	LRTARGETVEL : LREAL;
	LRTARGETPOS : LREAL;
	LRJERKACC : LREAL;
	LRJERKDEC : LREAL;
	LRJERKTIMEACC : LREAL;
	LRJERKTIMEDEC : LREAL;
	SCMAXPROFILEDATA : L_MB1P_IntProfileData;
	SCMINPROFILEDATA : L_MB1P_IntProfileData;
END_VAR
VAR_OUTPUT
	DWSTATE : DWORD;
END_VAR
VAR_IN_OUT
	SCPROFILEDATA : L_MB1P_ProfileData;
	SCPROFILEPARAMETER : L_MB1P_ProfileParameter;
END_VAR
END_METHOD

METHOD CALCPROFILE_20CB_AOGET0 : BOOL
VAR_INPUT
	LRSTARTACC : LREAL;
	LRSTARTVEL : LREAL;
	LRMAXACC : LREAL;
	LRMAXDEC : LREAL;
	LRMAXVEL : LREAL;
	LRTARGETACC : LREAL;
	LRTARGETVEL : LREAL;
	LRTARGETPOS : LREAL;
	LRJERKACC : LREAL;
	LRJERKDEC : LREAL;
	LRJERKTIMEACC : LREAL;
	LRJERKTIMEDEC : LREAL;
	T7 : LREAL;
END_VAR
VAR_IN_OUT
	SCPROFILEDATA : L_MB1P_ProfileData;
END_VAR
END_METHOD

METHOD CALCPROFILE_20CB_AOLT0 : BOOL
VAR_INPUT
	LRSTARTACC : LREAL;
	LRSTARTVEL : LREAL;
	LRMAXACC : LREAL;
	LRMAXDEC : LREAL;
	LRMAXVEL : LREAL;
	LRTARGETACC : LREAL;
	LRTARGETVEL : LREAL;
	LRTARGETPOS : LREAL;
	LRJERKACC : LREAL;
	LRJERKDEC : LREAL;
	LRJERKTIMEACC : LREAL;
	LRJERKTIMEDEC : LREAL;
	T7 : LREAL;
END_VAR
VAR_IN_OUT
	SCPROFILEDATA : L_MB1P_ProfileData;
END_VAR
END_METHOD

METHOD CALCPROFILE_20CBAOGET0_SEARCHTIMES : BOOL
VAR_INPUT
	LRSTARTACC : LREAL;
	LRSTARTVEL : LREAL;
	LRMAXACC : LREAL;
	LRMAXDEC : LREAL;
	LRMAXVEL : LREAL;
	LRTARGETACC : LREAL;
	LRTARGETVEL : LREAL;
	LRTARGETPOS : LREAL;
	LRJERKACC : LREAL;
	LRJERKDEC : LREAL;
	LRJERKTIMEACC : LREAL;
	LRJERKTIMEDEC : LREAL;
	T7_MINVALUE : LREAL;
	T7_MAXVALUE : LREAL;
END_VAR
VAR_OUTPUT
	T7 : LREAL;
END_VAR
END_METHOD

METHOD CALCPROFILE_20CBAOLT0_SEARCHTIMES : BOOL
VAR_INPUT
	LRSTARTACC : LREAL;
	LRSTARTVEL : LREAL;
	LRMAXACC : LREAL;
	LRMAXDEC : LREAL;
	LRMAXVEL : LREAL;
	LRTARGETACC : LREAL;
	LRTARGETVEL : LREAL;
	LRTARGETPOS : LREAL;
	LRJERKACC : LREAL;
	LRJERKDEC : LREAL;
	LRJERKTIMEACC : LREAL;
	LRJERKTIMEDEC : LREAL;
	T7_MINVALUE : LREAL;
	T7_MAXVALUE : LREAL;
END_VAR
VAR_OUTPUT
	T7 : LREAL;
END_VAR
END_METHOD

METHOD CALCPROFILE_20D0 : BOOL
VAR_INPUT
	LRSTARTACC : LREAL;
	LRSTARTVEL : LREAL;
	LRMAXACC : LREAL;
	LRMAXDEC : LREAL;
	LRMAXVEL : LREAL;
	LRTARGETACC : LREAL;
	LRTARGETVEL : LREAL;
	LRTARGETPOS : LREAL;
	LRJERKACC : LREAL;
	LRJERKDEC : LREAL;
	LRJERKTIMEACC : LREAL;
	LRJERKTIMEDEC : LREAL;
	SCMAXPROFILEDATA : L_MB1P_IntProfileData;
	SCMINPROFILEDATA : L_MB1P_IntProfileData;
END_VAR
VAR_OUTPUT
	DWSTATE : DWORD;
END_VAR
VAR_IN_OUT
	SCPROFILEDATA : L_MB1P_ProfileData;
	SCPROFILEPARAMETER : L_MB1P_ProfileParameter;
END_VAR
END_METHOD

METHOD CALCPROFILE_20D0_SEARCHTIMEST5T7 : BOOL
VAR_INPUT
	LRSTARTACC : LREAL;
	LRSTARTVEL : LREAL;
	LRMAXACC : LREAL;
	LRMAXDEC : LREAL;
	LRMAXVEL : LREAL;
	LRTARGETACC : LREAL;
	LRTARGETVEL : LREAL;
	LRTARGETPOS : LREAL;
	LRJERKACC : LREAL;
	LRJERKDEC : LREAL;
	LRJERKTIMEACC : LREAL;
	LRJERKTIMEDEC : LREAL;
	T5_STARTVALUE : LREAL;
	T7_STARTVALUE : LREAL;
END_VAR
VAR_OUTPUT
	T5 : LREAL;
	T7 : LREAL;
END_VAR
END_METHOD

METHOD CALCPROFILE_20D0_A0LTAMAXT5T7 : BOOL
VAR_INPUT
	LRSTARTACC : LREAL;
	LRSTARTVEL : LREAL;
	LRMAXACC : LREAL;
	LRMAXDEC : LREAL;
	LRMAXVEL : LREAL;
	LRTARGETACC : LREAL;
	LRTARGETVEL : LREAL;
	LRTARGETPOS : LREAL;
	LRJERKACC : LREAL;
	LRJERKDEC : LREAL;
	LRJERKTIMEACC : LREAL;
	LRJERKTIMEDEC : LREAL;
	T5 : LREAL;
	T7 : LREAL;
END_VAR
VAR_IN_OUT
	SCPROFILEDATA : L_MB1P_ProfileData;
END_VAR
END_METHOD

METHOD CALCPROFILE_20D1 : BOOL
VAR_INPUT
	LRSTARTACC : LREAL;
	LRSTARTVEL : LREAL;
	LRMAXACC : LREAL;
	LRMAXDEC : LREAL;
	LRMAXVEL : LREAL;
	LRTARGETACC : LREAL;
	LRTARGETVEL : LREAL;
	LRTARGETPOS : LREAL;
	LRJERKACC : LREAL;
	LRJERKDEC : LREAL;
	LRJERKTIMEACC : LREAL;
	LRJERKTIMEDEC : LREAL;
	SCMAXPROFILEDATA : L_MB1P_IntProfileData;
	SCMINPROFILEDATA : L_MB1P_IntProfileData;
END_VAR
VAR_OUTPUT
	DWSTATE : DWORD;
END_VAR
VAR_IN_OUT
	SCPROFILEDATA : L_MB1P_ProfileData;
	SCPROFILEPARAMETER : L_MB1P_ProfileParameter;
END_VAR
END_METHOD

METHOD CALCPROFILE_20D1_AOGET0 : BOOL
VAR_INPUT
	LRSTARTACC : LREAL;
	LRSTARTVEL : LREAL;
	LRMAXACC : LREAL;
	LRMAXDEC : LREAL;
	LRMAXVEL : LREAL;
	LRTARGETACC : LREAL;
	LRTARGETVEL : LREAL;
	LRTARGETPOS : LREAL;
	LRJERKACC : LREAL;
	LRJERKDEC : LREAL;
	LRJERKTIMEACC : LREAL;
	LRJERKTIMEDEC : LREAL;
	T7 : LREAL;
END_VAR
VAR_IN_OUT
	SCPROFILEDATA : L_MB1P_ProfileData;
END_VAR
END_METHOD

METHOD CALCPROFILE_20D1_AOLT0 : BOOL
VAR_INPUT
	LRSTARTACC : LREAL;
	LRSTARTVEL : LREAL;
	LRMAXACC : LREAL;
	LRMAXDEC : LREAL;
	LRMAXVEL : LREAL;
	LRTARGETACC : LREAL;
	LRTARGETVEL : LREAL;
	LRTARGETPOS : LREAL;
	LRJERKACC : LREAL;
	LRJERKDEC : LREAL;
	LRJERKTIMEACC : LREAL;
	LRJERKTIMEDEC : LREAL;
	T7 : LREAL;
END_VAR
VAR_IN_OUT
	SCPROFILEDATA : L_MB1P_ProfileData;
END_VAR
END_METHOD

METHOD CALCPROFILE_20D1AOGET0_SEARCHTIMES : BOOL
VAR_INPUT
	LRSTARTACC : LREAL;
	LRSTARTVEL : LREAL;
	LRMAXACC : LREAL;
	LRMAXDEC : LREAL;
	LRMAXVEL : LREAL;
	LRTARGETACC : LREAL;
	LRTARGETVEL : LREAL;
	LRTARGETPOS : LREAL;
	LRJERKACC : LREAL;
	LRJERKDEC : LREAL;
	LRJERKTIMEACC : LREAL;
	LRJERKTIMEDEC : LREAL;
	T7_STARTVALUE : LREAL;
END_VAR
VAR_OUTPUT
	T7 : LREAL;
END_VAR
END_METHOD

METHOD CALCPROFILE_20D1AOLT0_SEARCHTIMES : BOOL
VAR_INPUT
	LRSTARTACC : LREAL;
	LRSTARTVEL : LREAL;
	LRMAXACC : LREAL;
	LRMAXDEC : LREAL;
	LRMAXVEL : LREAL;
	LRTARGETACC : LREAL;
	LRTARGETVEL : LREAL;
	LRTARGETPOS : LREAL;
	LRJERKACC : LREAL;
	LRJERKDEC : LREAL;
	LRJERKTIMEACC : LREAL;
	LRJERKTIMEDEC : LREAL;
	T7_STARTVALUE : LREAL;
END_VAR
VAR_OUTPUT
	T7 : LREAL;
END_VAR
END_METHOD

METHOD CALCPROFILE_20DA : BOOL
VAR_INPUT
	LRSTARTACC : LREAL;
	LRSTARTVEL : LREAL;
	LRMAXACC : LREAL;
	LRMAXDEC : LREAL;
	LRMAXVEL : LREAL;
	LRTARGETACC : LREAL;
	LRTARGETVEL : LREAL;
	LRTARGETPOS : LREAL;
	LRJERKACC : LREAL;
	LRJERKDEC : LREAL;
	LRJERKTIMEACC : LREAL;
	LRJERKTIMEDEC : LREAL;
	SCMAXPROFILEDATA : L_MB1P_IntProfileData;
	SCMINPROFILEDATA : L_MB1P_IntProfileData;
END_VAR
VAR_OUTPUT
	DWSTATE : DWORD;
END_VAR
VAR_IN_OUT
	SCPROFILEDATA : L_MB1P_ProfileData;
	SCPROFILEPARAMETER : L_MB1P_ProfileParameter;
END_VAR
END_METHOD

METHOD CALCPROFILE_20DA_AELT0 : BOOL
VAR_INPUT
	LRSTARTACC : LREAL;
	LRSTARTVEL : LREAL;
	LRMAXACC : LREAL;
	LRMAXDEC : LREAL;
	LRMAXVEL : LREAL;
	LRTARGETACC : LREAL;
	LRTARGETVEL : LREAL;
	LRTARGETPOS : LREAL;
	LRJERKACC : LREAL;
	LRJERKDEC : LREAL;
	LRJERKTIMEACC : LREAL;
	LRJERKTIMEDEC : LREAL;
	T7 : LREAL;
END_VAR
VAR_IN_OUT
	SCPROFILEDATA : L_MB1P_ProfileData;
END_VAR
END_METHOD

METHOD CALCPROFILE_20DAAELT0_SEARCHTIMES : BOOL
VAR_INPUT
	LRSTARTACC : LREAL;
	LRSTARTVEL : LREAL;
	LRMAXACC : LREAL;
	LRMAXDEC : LREAL;
	LRMAXVEL : LREAL;
	LRTARGETACC : LREAL;
	LRTARGETVEL : LREAL;
	LRTARGETPOS : LREAL;
	LRJERKACC : LREAL;
	LRJERKDEC : LREAL;
	LRJERKTIMEACC : LREAL;
	LRJERKTIMEDEC : LREAL;
	T7_MINVALUE : LREAL;
	T7_MAXVALUE : LREAL;
END_VAR
VAR_OUTPUT
	T7 : LREAL;
END_VAR
END_METHOD

METHOD CALCPROFILE_20DB : BOOL
VAR_INPUT
	LRSTARTACC : LREAL;
	LRSTARTVEL : LREAL;
	LRMAXACC : LREAL;
	LRMAXDEC : LREAL;
	LRMAXVEL : LREAL;
	LRTARGETACC : LREAL;
	LRTARGETVEL : LREAL;
	LRTARGETPOS : LREAL;
	LRJERKACC : LREAL;
	LRJERKDEC : LREAL;
	LRJERKTIMEACC : LREAL;
	LRJERKTIMEDEC : LREAL;
	SCMAXPROFILEDATA : L_MB1P_IntProfileData;
	SCMINPROFILEDATA : L_MB1P_IntProfileData;
END_VAR
VAR_OUTPUT
	DWSTATE : DWORD;
END_VAR
VAR_IN_OUT
	SCPROFILEDATA : L_MB1P_ProfileData;
	SCPROFILEPARAMETER : L_MB1P_ProfileParameter;
END_VAR
END_METHOD

METHOD CALCPROFILE_20DB_AOGET0 : BOOL
VAR_INPUT
	LRSTARTACC : LREAL;
	LRSTARTVEL : LREAL;
	LRMAXACC : LREAL;
	LRMAXDEC : LREAL;
	LRMAXVEL : LREAL;
	LRTARGETACC : LREAL;
	LRTARGETVEL : LREAL;
	LRTARGETPOS : LREAL;
	LRJERKACC : LREAL;
	LRJERKDEC : LREAL;
	LRJERKTIMEACC : LREAL;
	LRJERKTIMEDEC : LREAL;
	T7 : LREAL;
END_VAR
VAR_IN_OUT
	SCPROFILEDATA : L_MB1P_ProfileData;
END_VAR
END_METHOD

METHOD CALCPROFILE_20DB_AOLT0 : BOOL
VAR_INPUT
	LRSTARTACC : LREAL;
	LRSTARTVEL : LREAL;
	LRMAXACC : LREAL;
	LRMAXDEC : LREAL;
	LRMAXVEL : LREAL;
	LRTARGETACC : LREAL;
	LRTARGETVEL : LREAL;
	LRTARGETPOS : LREAL;
	LRJERKACC : LREAL;
	LRJERKDEC : LREAL;
	LRJERKTIMEACC : LREAL;
	LRJERKTIMEDEC : LREAL;
	T7 : LREAL;
END_VAR
VAR_IN_OUT
	SCPROFILEDATA : L_MB1P_ProfileData;
END_VAR
END_METHOD

METHOD CALCPROFILE_20DBAOGET0_SEARCHTIMES : BOOL
VAR_INPUT
	LRSTARTACC : LREAL;
	LRSTARTVEL : LREAL;
	LRMAXACC : LREAL;
	LRMAXDEC : LREAL;
	LRMAXVEL : LREAL;
	LRTARGETACC : LREAL;
	LRTARGETVEL : LREAL;
	LRTARGETPOS : LREAL;
	LRJERKACC : LREAL;
	LRJERKDEC : LREAL;
	LRJERKTIMEACC : LREAL;
	LRJERKTIMEDEC : LREAL;
	T7_MINVALUE : LREAL;
	T7_MAXVALUE : LREAL;
END_VAR
VAR_OUTPUT
	T7 : LREAL;
END_VAR
END_METHOD

METHOD CALCPROFILE_20DBAOLT0_SEARCHTIMES : BOOL
VAR_INPUT
	LRSTARTACC : LREAL;
	LRSTARTVEL : LREAL;
	LRMAXACC : LREAL;
	LRMAXDEC : LREAL;
	LRMAXVEL : LREAL;
	LRTARGETACC : LREAL;
	LRTARGETVEL : LREAL;
	LRTARGETPOS : LREAL;
	LRJERKACC : LREAL;
	LRJERKDEC : LREAL;
	LRJERKTIMEACC : LREAL;
	LRJERKTIMEDEC : LREAL;
	T7_MINVALUE : LREAL;
	T7_MAXVALUE : LREAL;
END_VAR
VAR_OUTPUT
	T7 : LREAL;
END_VAR
END_METHOD

METHOD CALCPROFILE_30A0 : BOOL
VAR_INPUT
	LRSTARTACC : LREAL;
	LRSTARTVEL : LREAL;
	LRMAXACC : LREAL;
	LRMAXDEC : LREAL;
	LRMAXVEL : LREAL;
	LRTARGETACC : LREAL;
	LRTARGETVEL : LREAL;
	LRTARGETPOS : LREAL;
	LRJERKACC : LREAL;
	LRJERKDEC : LREAL;
	LRJERKTIMEACC : LREAL;
	LRJERKTIMEDEC : LREAL;
END_VAR
VAR_OUTPUT
	DWSTATE : DWORD;
END_VAR
VAR_IN_OUT
	SCPROFILEDATA : L_MB1P_ProfileData;
	SCPROFILEPARAMETER : L_MB1P_ProfileParameter;
END_VAR
END_METHOD

METHOD CALCPROFILE_30A0_A0GTAMAX : BOOL
VAR_INPUT
	LRSTARTACC : LREAL;
	LRSTARTVEL : LREAL;
	LRMAXACC : LREAL;
	LRMAXDEC : LREAL;
	LRMAXVEL : LREAL;
	LRTARGETACC : LREAL;
	LRTARGETVEL : LREAL;
	LRTARGETPOS : LREAL;
	LRJERKACC : LREAL;
	LRJERKDEC : LREAL;
	LRJERKTIMEACC : LREAL;
	LRJERKTIMEDEC : LREAL;
END_VAR
VAR_IN_OUT
	SCPROFILEDATA : L_MB1P_ProfileData;
END_VAR
END_METHOD

METHOD CALCPROFILE_30A0_A0LTAMAX : BOOL
VAR_INPUT
	LRSTARTACC : LREAL;
	LRSTARTVEL : LREAL;
	LRMAXACC : LREAL;
	LRMAXDEC : LREAL;
	LRMAXVEL : LREAL;
	LRTARGETACC : LREAL;
	LRTARGETVEL : LREAL;
	LRTARGETPOS : LREAL;
	LRJERKACC : LREAL;
	LRJERKDEC : LREAL;
	LRJERKTIMEACC : LREAL;
	LRJERKTIMEDEC : LREAL;
END_VAR
VAR_IN_OUT
	SCPROFILEDATA : L_MB1P_ProfileData;
END_VAR
END_METHOD

METHOD CALCPROFILE_30B0 : BOOL
VAR_INPUT
	LRSTARTACC : LREAL;
	LRSTARTVEL : LREAL;
	LRMAXACC : LREAL;
	LRMAXDEC : LREAL;
	LRMAXVEL : LREAL;
	LRTARGETACC : LREAL;
	LRTARGETVEL : LREAL;
	LRTARGETPOS : LREAL;
	LRJERKACC : LREAL;
	LRJERKDEC : LREAL;
	LRJERKTIMEACC : LREAL;
	LRJERKTIMEDEC : LREAL;
END_VAR
VAR_OUTPUT
	DWSTATE : DWORD;
END_VAR
VAR_IN_OUT
	SCPROFILEDATA : L_MB1P_ProfileData;
	SCPROFILEPARAMETER : L_MB1P_ProfileParameter;
END_VAR
END_METHOD

METHOD CALCPROFILE_30B0_A0GTAMAXT51 : BOOL
VAR_INPUT
	LRSTARTACC : LREAL;
	LRSTARTVEL : LREAL;
	LRMAXACC : LREAL;
	LRMAXDEC : LREAL;
	LRMAXVEL : LREAL;
	LRTARGETACC : LREAL;
	LRTARGETVEL : LREAL;
	LRTARGETPOS : LREAL;
	LRJERKACC : LREAL;
	LRJERKDEC : LREAL;
	LRJERKTIMEACC : LREAL;
	LRJERKTIMEDEC : LREAL;
END_VAR
VAR_IN_OUT
	SCPROFILEDATA : L_MB1P_ProfileData;
END_VAR
END_METHOD

METHOD CALCPROFILE_30B0_A0GTAMAXT52 : BOOL
VAR_INPUT
	LRSTARTACC : LREAL;
	LRSTARTVEL : LREAL;
	LRMAXACC : LREAL;
	LRMAXDEC : LREAL;
	LRMAXVEL : LREAL;
	LRTARGETACC : LREAL;
	LRTARGETVEL : LREAL;
	LRTARGETPOS : LREAL;
	LRJERKACC : LREAL;
	LRJERKDEC : LREAL;
	LRJERKTIMEACC : LREAL;
	LRJERKTIMEDEC : LREAL;
END_VAR
VAR_IN_OUT
	SCPROFILEDATA : L_MB1P_ProfileData;
END_VAR
END_METHOD

METHOD CALCPROFILE_30B0_A0LTAMAXT51 : BOOL
VAR_INPUT
	LRSTARTACC : LREAL;
	LRSTARTVEL : LREAL;
	LRMAXACC : LREAL;
	LRMAXDEC : LREAL;
	LRMAXVEL : LREAL;
	LRTARGETACC : LREAL;
	LRTARGETVEL : LREAL;
	LRTARGETPOS : LREAL;
	LRJERKACC : LREAL;
	LRJERKDEC : LREAL;
	LRJERKTIMEACC : LREAL;
	LRJERKTIMEDEC : LREAL;
END_VAR
VAR_IN_OUT
	SCPROFILEDATA : L_MB1P_ProfileData;
END_VAR
END_METHOD

METHOD CALCPROFILE_30B0_A0LTAMAXT52 : BOOL
VAR_INPUT
	LRSTARTACC : LREAL;
	LRSTARTVEL : LREAL;
	LRMAXACC : LREAL;
	LRMAXDEC : LREAL;
	LRMAXVEL : LREAL;
	LRTARGETACC : LREAL;
	LRTARGETVEL : LREAL;
	LRTARGETPOS : LREAL;
	LRJERKACC : LREAL;
	LRJERKDEC : LREAL;
	LRJERKTIMEACC : LREAL;
	LRJERKTIMEDEC : LREAL;
END_VAR
VAR_IN_OUT
	SCPROFILEDATA : L_MB1P_ProfileData;
END_VAR
END_METHOD

METHOD CALCPROFILE_30C0 : BOOL
VAR_INPUT
	LRSTARTACC : LREAL;
	LRSTARTVEL : LREAL;
	LRMAXACC : LREAL;
	LRMAXDEC : LREAL;
	LRMAXVEL : LREAL;
	LRTARGETACC : LREAL;
	LRTARGETVEL : LREAL;
	LRTARGETPOS : LREAL;
	LRJERKACC : LREAL;
	LRJERKDEC : LREAL;
	LRJERKTIMEACC : LREAL;
	LRJERKTIMEDEC : LREAL;
END_VAR
VAR_OUTPUT
	DWSTATE : DWORD;
END_VAR
VAR_IN_OUT
	SCPROFILEDATA : L_MB1P_ProfileData;
	SCPROFILEPARAMETER : L_MB1P_ProfileParameter;
END_VAR
END_METHOD

METHOD CALCPROFILE_30C0_A0GTAMAXT31 : BOOL
VAR_INPUT
	LRSTARTACC : LREAL;
	LRSTARTVEL : LREAL;
	LRMAXACC : LREAL;
	LRMAXDEC : LREAL;
	LRMAXVEL : LREAL;
	LRTARGETACC : LREAL;
	LRTARGETVEL : LREAL;
	LRTARGETPOS : LREAL;
	LRJERKACC : LREAL;
	LRJERKDEC : LREAL;
	LRJERKTIMEACC : LREAL;
	LRJERKTIMEDEC : LREAL;
END_VAR
VAR_IN_OUT
	SCPROFILEDATA : L_MB1P_ProfileData;
END_VAR
END_METHOD

METHOD CALCPROFILE_30C0_A0GTAMAXT32 : BOOL
VAR_INPUT
	LRSTARTACC : LREAL;
	LRSTARTVEL : LREAL;
	LRMAXACC : LREAL;
	LRMAXDEC : LREAL;
	LRMAXVEL : LREAL;
	LRTARGETACC : LREAL;
	LRTARGETVEL : LREAL;
	LRTARGETPOS : LREAL;
	LRJERKACC : LREAL;
	LRJERKDEC : LREAL;
	LRJERKTIMEACC : LREAL;
	LRJERKTIMEDEC : LREAL;
END_VAR
VAR_IN_OUT
	SCPROFILEDATA : L_MB1P_ProfileData;
END_VAR
END_METHOD

METHOD CALCPROFILE_30CB : BOOL
VAR_INPUT
	LRSTARTACC : LREAL;
	LRSTARTVEL : LREAL;
	LRMAXACC : LREAL;
	LRMAXDEC : LREAL;
	LRMAXVEL : LREAL;
	LRTARGETACC : LREAL;
	LRTARGETVEL : LREAL;
	LRTARGETPOS : LREAL;
	LRJERKACC : LREAL;
	LRJERKDEC : LREAL;
	LRJERKTIMEACC : LREAL;
	LRJERKTIMEDEC : LREAL;
	SCMAXPROFILEDATA : L_MB1P_IntProfileData;
	SCMINPROFILEDATA : L_MB1P_IntProfileData;
END_VAR
VAR_OUTPUT
	DWSTATE : DWORD;
END_VAR
VAR_IN_OUT
	SCPROFILEDATA : L_MB1P_ProfileData;
	SCPROFILEPARAMETER : L_MB1P_ProfileParameter;
END_VAR
END_METHOD

METHOD CALCPROFILE_30CB_PROFILEDATA : BOOL
VAR_INPUT
	LRSTARTACC : LREAL;
	LRSTARTVEL : LREAL;
	LRMAXACC : LREAL;
	LRMAXDEC : LREAL;
	LRMAXVEL : LREAL;
	LRTARGETACC : LREAL;
	LRTARGETVEL : LREAL;
	LRTARGETPOS : LREAL;
	LRJERKACC : LREAL;
	LRJERKDEC : LREAL;
	LRJERKTIMEACC : LREAL;
	LRJERKTIMEDEC : LREAL;
	T7 : LREAL;
END_VAR
VAR_IN_OUT
	SCPROFILEDATA : L_MB1P_ProfileData;
END_VAR
END_METHOD

METHOD CALCPROFILE_30CB_SEARCHTIMES : BOOL
VAR_INPUT
	LRSTARTACC : LREAL;
	LRSTARTVEL : LREAL;
	LRMAXACC : LREAL;
	LRMAXDEC : LREAL;
	LRMAXVEL : LREAL;
	LRTARGETACC : LREAL;
	LRTARGETVEL : LREAL;
	LRTARGETPOS : LREAL;
	LRJERKACC : LREAL;
	LRJERKDEC : LREAL;
	LRJERKTIMEACC : LREAL;
	LRJERKTIMEDEC : LREAL;
	T7_MINVALUE : LREAL;
	T7_MAXVALUE : LREAL;
END_VAR
VAR_OUTPUT
	T7 : LREAL;
END_VAR
END_METHOD

METHOD CALCPROFILE_30D0 : BOOL
VAR_INPUT
	LRSTARTACC : LREAL;
	LRSTARTVEL : LREAL;
	LRMAXACC : LREAL;
	LRMAXDEC : LREAL;
	LRMAXVEL : LREAL;
	LRTARGETACC : LREAL;
	LRTARGETVEL : LREAL;
	LRTARGETPOS : LREAL;
	LRJERKACC : LREAL;
	LRJERKDEC : LREAL;
	LRJERKTIMEACC : LREAL;
	LRJERKTIMEDEC : LREAL;
END_VAR
VAR_OUTPUT
	DWSTATE : DWORD;
END_VAR
VAR_IN_OUT
	SCPROFILEDATA : L_MB1P_ProfileData;
	SCPROFILEPARAMETER : L_MB1P_ProfileParameter;
END_VAR
END_METHOD

METHOD CALCPROFILE_30D0_A0GTAMAXT31T51 : BOOL
VAR_INPUT
	LRSTARTACC : LREAL;
	LRSTARTVEL : LREAL;
	LRMAXACC : LREAL;
	LRMAXDEC : LREAL;
	LRMAXVEL : LREAL;
	LRTARGETACC : LREAL;
	LRTARGETVEL : LREAL;
	LRTARGETPOS : LREAL;
	LRJERKACC : LREAL;
	LRJERKDEC : LREAL;
	LRJERKTIMEACC : LREAL;
	LRJERKTIMEDEC : LREAL;
END_VAR
VAR_IN_OUT
	SCPROFILEDATA : L_MB1P_ProfileData;
END_VAR
END_METHOD

METHOD CALCPROFILE_30D0_A0GTAMAXT31T52 : BOOL
VAR_INPUT
	LRSTARTACC : LREAL;
	LRSTARTVEL : LREAL;
	LRMAXACC : LREAL;
	LRMAXDEC : LREAL;
	LRMAXVEL : LREAL;
	LRTARGETACC : LREAL;
	LRTARGETVEL : LREAL;
	LRTARGETPOS : LREAL;
	LRJERKACC : LREAL;
	LRJERKDEC : LREAL;
	LRJERKTIMEACC : LREAL;
	LRJERKTIMEDEC : LREAL;
END_VAR
VAR_IN_OUT
	SCPROFILEDATA : L_MB1P_ProfileData;
END_VAR
END_METHOD

METHOD CALCPROFILE_30D0_A0GTAMAXT32T51 : BOOL
VAR_INPUT
	LRSTARTACC : LREAL;
	LRSTARTVEL : LREAL;
	LRMAXACC : LREAL;
	LRMAXDEC : LREAL;
	LRMAXVEL : LREAL;
	LRTARGETACC : LREAL;
	LRTARGETVEL : LREAL;
	LRTARGETPOS : LREAL;
	LRJERKACC : LREAL;
	LRJERKDEC : LREAL;
	LRJERKTIMEACC : LREAL;
	LRJERKTIMEDEC : LREAL;
END_VAR
VAR_IN_OUT
	SCPROFILEDATA : L_MB1P_ProfileData;
END_VAR
END_METHOD

METHOD CALCPROFILE_30D0_A0GTAMAXT32T52 : BOOL
VAR_INPUT
	LRSTARTACC : LREAL;
	LRSTARTVEL : LREAL;
	LRMAXACC : LREAL;
	LRMAXDEC : LREAL;
	LRMAXVEL : LREAL;
	LRTARGETACC : LREAL;
	LRTARGETVEL : LREAL;
	LRTARGETPOS : LREAL;
	LRJERKACC : LREAL;
	LRJERKDEC : LREAL;
	LRJERKTIMEACC : LREAL;
	LRJERKTIMEDEC : LREAL;
END_VAR
VAR_IN_OUT
	SCPROFILEDATA : L_MB1P_ProfileData;
END_VAR
END_METHOD

METHOD CALCPROFILE_30D1 : BOOL
VAR_INPUT
	LRSTARTACC : LREAL;
	LRSTARTVEL : LREAL;
	LRMAXACC : LREAL;
	LRMAXDEC : LREAL;
	LRMAXVEL : LREAL;
	LRTARGETACC : LREAL;
	LRTARGETVEL : LREAL;
	LRTARGETPOS : LREAL;
	LRJERKACC : LREAL;
	LRJERKDEC : LREAL;
	LRJERKTIMEACC : LREAL;
	LRJERKTIMEDEC : LREAL;
	SCMAXPROFILEDATA : L_MB1P_IntProfileData;
	SCMINPROFILEDATA : L_MB1P_IntProfileData;
END_VAR
VAR_OUTPUT
	DWSTATE : DWORD;
END_VAR
VAR_IN_OUT
	SCPROFILEDATA : L_MB1P_ProfileData;
	SCPROFILEPARAMETER : L_MB1P_ProfileParameter;
END_VAR
END_METHOD

METHOD CALCPROFILE_30D1_PROFILEDATA : BOOL
VAR_INPUT
	LRSTARTACC : LREAL;
	LRSTARTVEL : LREAL;
	LRMAXACC : LREAL;
	LRMAXDEC : LREAL;
	LRMAXVEL : LREAL;
	LRTARGETACC : LREAL;
	LRTARGETVEL : LREAL;
	LRTARGETPOS : LREAL;
	LRJERKACC : LREAL;
	LRJERKDEC : LREAL;
	LRJERKTIMEACC : LREAL;
	LRJERKTIMEDEC : LREAL;
	T7 : LREAL;
END_VAR
VAR_IN_OUT
	SCPROFILEDATA : L_MB1P_ProfileData;
END_VAR
END_METHOD

METHOD CALCPROFILE_30D1_SEARCHTIMES : BOOL
VAR_INPUT
	LRSTARTACC : LREAL;
	LRSTARTVEL : LREAL;
	LRMAXACC : LREAL;
	LRMAXDEC : LREAL;
	LRMAXVEL : LREAL;
	LRTARGETACC : LREAL;
	LRTARGETVEL : LREAL;
	LRTARGETPOS : LREAL;
	LRJERKACC : LREAL;
	LRJERKDEC : LREAL;
	LRJERKTIMEACC : LREAL;
	LRJERKTIMEDEC : LREAL;
	T7_MINVALUE : LREAL;
	T7_MAXVALUE : LREAL;
END_VAR
VAR_OUTPUT
	T7 : LREAL;
END_VAR
END_METHOD

METHOD CALCPROFILE_30DB : BOOL
VAR_INPUT
	LRSTARTACC : LREAL;
	LRSTARTVEL : LREAL;
	LRMAXACC : LREAL;
	LRMAXDEC : LREAL;
	LRMAXVEL : LREAL;
	LRTARGETACC : LREAL;
	LRTARGETVEL : LREAL;
	LRTARGETPOS : LREAL;
	LRJERKACC : LREAL;
	LRJERKDEC : LREAL;
	LRJERKTIMEACC : LREAL;
	LRJERKTIMEDEC : LREAL;
	SCMAXPROFILEDATA : L_MB1P_IntProfileData;
	SCMINPROFILEDATA : L_MB1P_IntProfileData;
END_VAR
VAR_OUTPUT
	DWSTATE : DWORD;
END_VAR
VAR_IN_OUT
	SCPROFILEDATA : L_MB1P_ProfileData;
	SCPROFILEPARAMETER : L_MB1P_ProfileParameter;
END_VAR
END_METHOD

METHOD CALCPROFILE_30DB_PROFILEDATA : BOOL
VAR_INPUT
	LRSTARTACC : LREAL;
	LRSTARTVEL : LREAL;
	LRMAXACC : LREAL;
	LRMAXDEC : LREAL;
	LRMAXVEL : LREAL;
	LRTARGETACC : LREAL;
	LRTARGETVEL : LREAL;
	LRTARGETPOS : LREAL;
	LRJERKACC : LREAL;
	LRJERKDEC : LREAL;
	LRJERKTIMEACC : LREAL;
	LRJERKTIMEDEC : LREAL;
	T7 : LREAL;
END_VAR
VAR_IN_OUT
	SCPROFILEDATA : L_MB1P_ProfileData;
END_VAR
END_METHOD

METHOD CALCPROFILE_30DB_SEARCHTIMES : BOOL
VAR_INPUT
	LRSTARTACC : LREAL;
	LRSTARTVEL : LREAL;
	LRMAXACC : LREAL;
	LRMAXDEC : LREAL;
	LRMAXVEL : LREAL;
	LRTARGETACC : LREAL;
	LRTARGETVEL : LREAL;
	LRTARGETPOS : LREAL;
	LRJERKACC : LREAL;
	LRJERKDEC : LREAL;
	LRJERKTIMEACC : LREAL;
	LRJERKTIMEDEC : LREAL;
	T7_MINVALUE : LREAL;
	T7_MAXVALUE : LREAL;
END_VAR
VAR_OUTPUT
	T7 : LREAL;
END_VAR
END_METHOD

METHOD CALCPROFILE_40A0 : BOOL
VAR_INPUT
	LRSTARTACC : LREAL;
	LRSTARTVEL : LREAL;
	LRMAXACC : LREAL;
	LRMAXDEC : LREAL;
	LRMAXVEL : LREAL;
	LRTARGETACC : LREAL;
	LRTARGETVEL : LREAL;
	LRTARGETPOS : LREAL;
	LRJERKACC : LREAL;
	LRJERKDEC : LREAL;
	LRJERKTIMEACC : LREAL;
	LRJERKTIMEDEC : LREAL;
END_VAR
VAR_OUTPUT
	DWSTATE : DWORD;
END_VAR
VAR_IN_OUT
	SCPROFILEDATA : L_MB1P_ProfileData;
	SCPROFILEPARAMETER : L_MB1P_ProfileParameter;
END_VAR
END_METHOD

METHOD CALCPROFILE_40A0_A0GTAMAX : BOOL
VAR_INPUT
	LRSTARTACC : LREAL;
	LRSTARTVEL : LREAL;
	LRMAXACC : LREAL;
	LRMAXDEC : LREAL;
	LRMAXVEL : LREAL;
	LRTARGETACC : LREAL;
	LRTARGETVEL : LREAL;
	LRTARGETPOS : LREAL;
	LRJERKACC : LREAL;
	LRJERKDEC : LREAL;
	LRJERKTIMEACC : LREAL;
	LRJERKTIMEDEC : LREAL;
END_VAR
VAR_IN_OUT
	SCPROFILEDATA : L_MB1P_ProfileData;
END_VAR
END_METHOD

METHOD CALCPROFILE_40A0_A0LTAMAX : BOOL
VAR_INPUT
	LRSTARTACC : LREAL;
	LRSTARTVEL : LREAL;
	LRMAXACC : LREAL;
	LRMAXDEC : LREAL;
	LRMAXVEL : LREAL;
	LRTARGETACC : LREAL;
	LRTARGETVEL : LREAL;
	LRTARGETPOS : LREAL;
	LRJERKACC : LREAL;
	LRJERKDEC : LREAL;
	LRJERKTIMEACC : LREAL;
	LRJERKTIMEDEC : LREAL;
END_VAR
VAR_IN_OUT
	SCPROFILEDATA : L_MB1P_ProfileData;
END_VAR
END_METHOD

METHOD CALCPROFILE_40B0 : BOOL
VAR_INPUT
	LRSTARTACC : LREAL;
	LRSTARTVEL : LREAL;
	LRMAXACC : LREAL;
	LRMAXDEC : LREAL;
	LRMAXVEL : LREAL;
	LRTARGETACC : LREAL;
	LRTARGETVEL : LREAL;
	LRTARGETPOS : LREAL;
	LRJERKACC : LREAL;
	LRJERKDEC : LREAL;
	LRJERKTIMEACC : LREAL;
	LRJERKTIMEDEC : LREAL;
END_VAR
VAR_OUTPUT
	DWSTATE : DWORD;
END_VAR
VAR_IN_OUT
	SCPROFILEDATA : L_MB1P_ProfileData;
	SCPROFILEPARAMETER : L_MB1P_ProfileParameter;
END_VAR
END_METHOD

METHOD CALCPROFILE_40C0 : BOOL
VAR_INPUT
	LRSTARTACC : LREAL;
	LRSTARTVEL : LREAL;
	LRMAXACC : LREAL;
	LRMAXDEC : LREAL;
	LRMAXVEL : LREAL;
	LRTARGETACC : LREAL;
	LRTARGETVEL : LREAL;
	LRTARGETPOS : LREAL;
	LRJERKACC : LREAL;
	LRJERKDEC : LREAL;
	LRJERKTIMEACC : LREAL;
	LRJERKTIMEDEC : LREAL;
END_VAR
VAR_OUTPUT
	DWSTATE : DWORD;
END_VAR
VAR_IN_OUT
	SCPROFILEDATA : L_MB1P_ProfileData;
	SCPROFILEPARAMETER : L_MB1P_ProfileParameter;
END_VAR
END_METHOD

METHOD CALCPROFILE_40C0_A0LTAMAXT31 : BOOL
VAR_INPUT
	LRSTARTACC : LREAL;
	LRSTARTVEL : LREAL;
	LRMAXACC : LREAL;
	LRMAXDEC : LREAL;
	LRMAXVEL : LREAL;
	LRTARGETACC : LREAL;
	LRTARGETVEL : LREAL;
	LRTARGETPOS : LREAL;
	LRJERKACC : LREAL;
	LRJERKDEC : LREAL;
	LRJERKTIMEACC : LREAL;
	LRJERKTIMEDEC : LREAL;
END_VAR
VAR_IN_OUT
	SCPROFILEDATA : L_MB1P_ProfileData;
END_VAR
END_METHOD

METHOD CALCPROFILE_40C0_A0LTAMAXT32 : BOOL
VAR_INPUT
	LRSTARTACC : LREAL;
	LRSTARTVEL : LREAL;
	LRMAXACC : LREAL;
	LRMAXDEC : LREAL;
	LRMAXVEL : LREAL;
	LRTARGETACC : LREAL;
	LRTARGETVEL : LREAL;
	LRTARGETPOS : LREAL;
	LRJERKACC : LREAL;
	LRJERKDEC : LREAL;
	LRJERKTIMEACC : LREAL;
	LRJERKTIMEDEC : LREAL;
END_VAR
VAR_IN_OUT
	SCPROFILEDATA : L_MB1P_ProfileData;
END_VAR
END_METHOD

METHOD CALCPROFILE_40D0 : BOOL
VAR_INPUT
	LRSTARTACC : LREAL;
	LRSTARTVEL : LREAL;
	LRMAXACC : LREAL;
	LRMAXDEC : LREAL;
	LRMAXVEL : LREAL;
	LRTARGETACC : LREAL;
	LRTARGETVEL : LREAL;
	LRTARGETPOS : LREAL;
	LRJERKACC : LREAL;
	LRJERKDEC : LREAL;
	LRJERKTIMEACC : LREAL;
	LRJERKTIMEDEC : LREAL;
END_VAR
VAR_OUTPUT
	DWSTATE : DWORD;
END_VAR
VAR_IN_OUT
	SCPROFILEDATA : L_MB1P_ProfileData;
	SCPROFILEPARAMETER : L_MB1P_ProfileParameter;
END_VAR
END_METHOD

METHOD CALCPROFILE_40E0 : BOOL
VAR_INPUT
	LRSTARTACC : LREAL;
	LRSTARTVEL : LREAL;
	LRMAXACC : LREAL;
	LRMAXDEC : LREAL;
	LRMAXVEL : LREAL;
	LRTARGETACC : LREAL;
	LRTARGETVEL : LREAL;
	LRTARGETPOS : LREAL;
	LRJERKACC : LREAL;
	LRJERKDEC : LREAL;
	LRJERKTIMEACC : LREAL;
	LRJERKTIMEDEC : LREAL;
END_VAR
VAR_OUTPUT
	DWSTATE : DWORD;
END_VAR
VAR_IN_OUT
	SCPROFILEDATA : L_MB1P_ProfileData;
	SCPROFILEPARAMETER : L_MB1P_ProfileParameter;
END_VAR
END_METHOD

METHOD CALCPROFILE_40F0 : BOOL
VAR_INPUT
	LRSTARTACC : LREAL;
	LRSTARTVEL : LREAL;
	LRMAXACC : LREAL;
	LRMAXDEC : LREAL;
	LRMAXVEL : LREAL;
	LRTARGETACC : LREAL;
	LRTARGETVEL : LREAL;
	LRTARGETPOS : LREAL;
	LRJERKACC : LREAL;
	LRJERKDEC : LREAL;
	LRJERKTIMEACC : LREAL;
	LRJERKTIMEDEC : LREAL;
END_VAR
VAR_OUTPUT
	DWSTATE : DWORD;
END_VAR
VAR_IN_OUT
	SCPROFILEDATA : L_MB1P_ProfileData;
	SCPROFILEPARAMETER : L_MB1P_ProfileParameter;
END_VAR
END_METHOD

METHOD CALCPROFILE_40F0_T51 : BOOL
VAR_INPUT
	LRSTARTACC : LREAL;
	LRSTARTVEL : LREAL;
	LRMAXACC : LREAL;
	LRMAXDEC : LREAL;
	LRMAXVEL : LREAL;
	LRTARGETACC : LREAL;
	LRTARGETVEL : LREAL;
	LRTARGETPOS : LREAL;
	LRJERKACC : LREAL;
	LRJERKDEC : LREAL;
	LRJERKTIMEACC : LREAL;
	LRJERKTIMEDEC : LREAL;
END_VAR
VAR_IN_OUT
	SCPROFILEDATA : L_MB1P_ProfileData;
END_VAR
END_METHOD

METHOD CALCPROFILE_40F0_T52 : BOOL
VAR_INPUT
	LRSTARTACC : LREAL;
	LRSTARTVEL : LREAL;
	LRMAXACC : LREAL;
	LRMAXDEC : LREAL;
	LRMAXVEL : LREAL;
	LRTARGETACC : LREAL;
	LRTARGETVEL : LREAL;
	LRTARGETPOS : LREAL;
	LRJERKACC : LREAL;
	LRJERKDEC : LREAL;
	LRJERKTIMEACC : LREAL;
	LRJERKTIMEDEC : LREAL;
END_VAR
VAR_IN_OUT
	SCPROFILEDATA : L_MB1P_ProfileData;
END_VAR
END_METHOD

METHOD CALCPROFILE_50A0 : BOOL
VAR_INPUT
	LRSTARTACC : LREAL;
	LRSTARTVEL : LREAL;
	LRMAXACC : LREAL;
	LRMAXDEC : LREAL;
	LRMAXVEL : LREAL;
	LRTARGETACC : LREAL;
	LRTARGETVEL : LREAL;
	LRTARGETPOS : LREAL;
	LRJERKACC : LREAL;
	LRJERKDEC : LREAL;
	LRJERKTIMEACC : LREAL;
	LRJERKTIMEDEC : LREAL;
END_VAR
VAR_OUTPUT
	DWSTATE : DWORD;
END_VAR
VAR_IN_OUT
	SCPROFILEDATA : L_MB1P_ProfileData;
	SCPROFILEPARAMETER : L_MB1P_ProfileParameter;
END_VAR
END_METHOD

METHOD CALCPROFILE_60A0 : BOOL
VAR_INPUT
	LRSTARTACC : LREAL;
	LRSTARTVEL : LREAL;
	LRMAXACC : LREAL;
	LRMAXDEC : LREAL;
	LRMAXVEL : LREAL;
	LRTARGETACC : LREAL;
	LRTARGETVEL : LREAL;
	LRTARGETPOS : LREAL;
	LRJERKACC : LREAL;
	LRJERKDEC : LREAL;
	LRJERKTIMEACC : LREAL;
	LRJERKTIMEDEC : LREAL;
END_VAR
VAR_OUTPUT
	DWSTATE : DWORD;
END_VAR
VAR_IN_OUT
	SCPROFILEDATA : L_MB1P_ProfileData;
	SCPROFILEPARAMETER : L_MB1P_ProfileParameter;
END_VAR
END_METHOD

METHOD CALCPROFILE_60A0_A0GTAMAX : BOOL
VAR_INPUT
	LRSTARTACC : LREAL;
	LRSTARTVEL : LREAL;
	LRMAXACC : LREAL;
	LRMAXDEC : LREAL;
	LRMAXVEL : LREAL;
	LRTARGETACC : LREAL;
	LRTARGETVEL : LREAL;
	LRTARGETPOS : LREAL;
	LRJERKACC : LREAL;
	LRJERKDEC : LREAL;
	LRJERKTIMEACC : LREAL;
	LRJERKTIMEDEC : LREAL;
END_VAR
VAR_IN_OUT
	SCPROFILEDATA : L_MB1P_ProfileData;
END_VAR
END_METHOD

METHOD CALCPROFILE_60A0_A0LTAMAX : BOOL
VAR_INPUT
	LRSTARTACC : LREAL;
	LRSTARTVEL : LREAL;
	LRMAXACC : LREAL;
	LRMAXDEC : LREAL;
	LRMAXVEL : LREAL;
	LRTARGETACC : LREAL;
	LRTARGETVEL : LREAL;
	LRTARGETPOS : LREAL;
	LRJERKACC : LREAL;
	LRJERKDEC : LREAL;
	LRJERKTIMEACC : LREAL;
	LRJERKTIMEDEC : LREAL;
END_VAR
VAR_IN_OUT
	SCPROFILEDATA : L_MB1P_ProfileData;
END_VAR
END_METHOD

METHOD CALCPROFILE_60B0 : BOOL
VAR_INPUT
	LRSTARTACC : LREAL;
	LRSTARTVEL : LREAL;
	LRMAXACC : LREAL;
	LRMAXDEC : LREAL;
	LRMAXVEL : LREAL;
	LRTARGETACC : LREAL;
	LRTARGETVEL : LREAL;
	LRTARGETPOS : LREAL;
	LRJERKACC : LREAL;
	LRJERKDEC : LREAL;
	LRJERKTIMEACC : LREAL;
	LRJERKTIMEDEC : LREAL;
END_VAR
VAR_OUTPUT
	DWSTATE : DWORD;
END_VAR
VAR_IN_OUT
	SCPROFILEDATA : L_MB1P_ProfileData;
	SCPROFILEPARAMETER : L_MB1P_ProfileParameter;
END_VAR
END_METHOD

METHOD CALCPROFILE_60B0_A0GTAMAX : BOOL
VAR_INPUT
	LRSTARTACC : LREAL;
	LRSTARTVEL : LREAL;
	LRMAXACC : LREAL;
	LRMAXDEC : LREAL;
	LRMAXVEL : LREAL;
	LRTARGETACC : LREAL;
	LRTARGETVEL : LREAL;
	LRTARGETPOS : LREAL;
	LRJERKACC : LREAL;
	LRJERKDEC : LREAL;
	LRJERKTIMEACC : LREAL;
	LRJERKTIMEDEC : LREAL;
END_VAR
VAR_IN_OUT
	SCPROFILEDATA : L_MB1P_ProfileData;
END_VAR
END_METHOD

METHOD CALCPROFILE_60B0_A0LTAMAX : BOOL
VAR_INPUT
	LRSTARTACC : LREAL;
	LRSTARTVEL : LREAL;
	LRMAXACC : LREAL;
	LRMAXDEC : LREAL;
	LRMAXVEL : LREAL;
	LRTARGETACC : LREAL;
	LRTARGETVEL : LREAL;
	LRTARGETPOS : LREAL;
	LRJERKACC : LREAL;
	LRJERKDEC : LREAL;
	LRJERKTIMEACC : LREAL;
	LRJERKTIMEDEC : LREAL;
END_VAR
VAR_IN_OUT
	SCPROFILEDATA : L_MB1P_ProfileData;
END_VAR
END_METHOD

METHOD CALCPROFILE_60C0 : BOOL
VAR_INPUT
	LRSTARTACC : LREAL;
	LRSTARTVEL : LREAL;
	LRMAXACC : LREAL;
	LRMAXDEC : LREAL;
	LRMAXVEL : LREAL;
	LRTARGETACC : LREAL;
	LRTARGETVEL : LREAL;
	LRTARGETPOS : LREAL;
	LRJERKACC : LREAL;
	LRJERKDEC : LREAL;
	LRJERKTIMEACC : LREAL;
	LRJERKTIMEDEC : LREAL;
END_VAR
VAR_OUTPUT
	DWSTATE : DWORD;
END_VAR
VAR_IN_OUT
	SCPROFILEDATA : L_MB1P_ProfileData;
	SCPROFILEPARAMETER : L_MB1P_ProfileParameter;
END_VAR
END_METHOD

METHOD CALCPROFILE_60D0 : BOOL
VAR_INPUT
	LRSTARTACC : LREAL;
	LRSTARTVEL : LREAL;
	LRMAXACC : LREAL;
	LRMAXDEC : LREAL;
	LRMAXVEL : LREAL;
	LRTARGETACC : LREAL;
	LRTARGETVEL : LREAL;
	LRTARGETPOS : LREAL;
	LRJERKACC : LREAL;
	LRJERKDEC : LREAL;
	LRJERKTIMEACC : LREAL;
	LRJERKTIMEDEC : LREAL;
END_VAR
VAR_OUTPUT
	DWSTATE : DWORD;
END_VAR
VAR_IN_OUT
	SCPROFILEDATA : L_MB1P_ProfileData;
	SCPROFILEPARAMETER : L_MB1P_ProfileParameter;
END_VAR
END_METHOD

METHOD CALCPROFILE_70A0 : BOOL
VAR_INPUT
	LRSTARTACC : LREAL;
	LRSTARTVEL : LREAL;
	LRMAXACC : LREAL;
	LRMAXDEC : LREAL;
	LRMAXVEL : LREAL;
	LRTARGETACC : LREAL;
	LRTARGETVEL : LREAL;
	LRTARGETPOS : LREAL;
	LRJERKACC : LREAL;
	LRJERKDEC : LREAL;
	LRJERKTIMEACC : LREAL;
	LRJERKTIMEDEC : LREAL;
	SCMAXPROFILEDATA : L_MB1P_IntProfileData;
	SCMINPROFILEDATA : L_MB1P_IntProfileData;
END_VAR
VAR_OUTPUT
	DWSTATE : DWORD;
END_VAR
VAR_IN_OUT
	SCPROFILEDATA : L_MB1P_ProfileData;
	SCPROFILEPARAMETER : L_MB1P_ProfileParameter;
END_VAR
END_METHOD

METHOD CALCPROFILE_70A0_SEARCHTIMEST5T7 : BOOL
VAR_INPUT
	LRSTARTACC : LREAL;
	LRSTARTVEL : LREAL;
	LRMAXACC : LREAL;
	LRMAXDEC : LREAL;
	LRMAXVEL : LREAL;
	LRTARGETACC : LREAL;
	LRTARGETVEL : LREAL;
	LRTARGETPOS : LREAL;
	LRJERKACC : LREAL;
	LRJERKDEC : LREAL;
	LRJERKTIMEACC : LREAL;
	LRJERKTIMEDEC : LREAL;
	T5_STARTVALUE : LREAL;
	T7_STARTVALUE : LREAL;
END_VAR
VAR_OUTPUT
	T5 : LREAL;
	T7 : LREAL;
END_VAR
END_METHOD

METHOD CALCPROFILE_70A0_A0LTAMAXT5T7 : BOOL
VAR_INPUT
	LRSTARTACC : LREAL;
	LRSTARTVEL : LREAL;
	LRMAXACC : LREAL;
	LRMAXDEC : LREAL;
	LRMAXVEL : LREAL;
	LRTARGETACC : LREAL;
	LRTARGETVEL : LREAL;
	LRTARGETPOS : LREAL;
	LRJERKACC : LREAL;
	LRJERKDEC : LREAL;
	LRJERKTIMEACC : LREAL;
	LRJERKTIMEDEC : LREAL;
	T5 : LREAL;
	T7 : LREAL;
END_VAR
VAR_OUTPUT
	A : ARRAY [1..4] OF LREAL;
END_VAR
VAR_IN_OUT
	SCPROFILEDATA : L_MB1P_ProfileData;
END_VAR
END_METHOD

METHOD CALCPROFILE_70B0 : BOOL
VAR_INPUT
	LRSTARTACC : LREAL;
	LRSTARTVEL : LREAL;
	LRMAXACC : LREAL;
	LRMAXDEC : LREAL;
	LRMAXVEL : LREAL;
	LRTARGETACC : LREAL;
	LRTARGETVEL : LREAL;
	LRTARGETPOS : LREAL;
	LRJERKACC : LREAL;
	LRJERKDEC : LREAL;
	LRJERKTIMEACC : LREAL;
	LRJERKTIMEDEC : LREAL;
	SCMAXPROFILEDATA : L_MB1P_IntProfileData;
	SCMINPROFILEDATA : L_MB1P_IntProfileData;
END_VAR
VAR_OUTPUT
	DWSTATE : DWORD;
END_VAR
VAR_IN_OUT
	SCPROFILEDATA : L_MB1P_ProfileData;
	SCPROFILEPARAMETER : L_MB1P_ProfileParameter;
END_VAR
END_METHOD

METHOD CALCPROFILE_70B0_SEARCHTIMEST5T7 : BOOL
VAR_INPUT
	LRSTARTACC : LREAL;
	LRSTARTVEL : LREAL;
	LRMAXACC : LREAL;
	LRMAXDEC : LREAL;
	LRMAXVEL : LREAL;
	LRTARGETACC : LREAL;
	LRTARGETVEL : LREAL;
	LRTARGETPOS : LREAL;
	LRJERKACC : LREAL;
	LRJERKDEC : LREAL;
	LRJERKTIMEACC : LREAL;
	LRJERKTIMEDEC : LREAL;
	T5_STARTVALUE : LREAL;
	T7_STARTVALUE : LREAL;
END_VAR
VAR_OUTPUT
	T5 : LREAL;
	T7 : LREAL;
END_VAR
END_METHOD

METHOD CALCPROFILE_70B0_A0LTAMAXT5T7 : BOOL
VAR_INPUT
	LRSTARTACC : LREAL;
	LRSTARTVEL : LREAL;
	LRMAXACC : LREAL;
	LRMAXDEC : LREAL;
	LRMAXVEL : LREAL;
	LRTARGETACC : LREAL;
	LRTARGETVEL : LREAL;
	LRTARGETPOS : LREAL;
	LRJERKACC : LREAL;
	LRJERKDEC : LREAL;
	LRJERKTIMEACC : LREAL;
	LRJERKTIMEDEC : LREAL;
	T5 : LREAL;
	T7 : LREAL;
END_VAR
VAR_OUTPUT
	A : ARRAY [1..4] OF LREAL;
END_VAR
VAR_IN_OUT
	SCPROFILEDATA : L_MB1P_ProfileData;
END_VAR
END_METHOD

METHOD CALCPROFILE_80A0 : BOOL
VAR_INPUT
	LRSTARTACC : LREAL;
	LRSTARTVEL : LREAL;
	LRMAXACC : LREAL;
	LRMAXDEC : LREAL;
	LRMAXVEL : LREAL;
	LRTARGETACC : LREAL;
	LRTARGETVEL : LREAL;
	LRTARGETPOS : LREAL;
	LRJERKACC : LREAL;
	LRJERKDEC : LREAL;
	LRJERKTIMEACC : LREAL;
	LRJERKTIMEDEC : LREAL;
	SCMAXPROFILEDATA : L_MB1P_IntProfileData;
	SCMINPROFILEDATA : L_MB1P_IntProfileData;
END_VAR
VAR_OUTPUT
	DWSTATE : DWORD;
END_VAR
VAR_IN_OUT
	SCPROFILEDATA : L_MB1P_ProfileData;
	SCPROFILEPARAMETER : L_MB1P_ProfileParameter;
END_VAR
END_METHOD

METHOD CALCPROFILE_80A0_A0GTAMAXT5T7 : BOOL
VAR_INPUT
	LRSTARTACC : LREAL;
	LRSTARTVEL : LREAL;
	LRMAXACC : LREAL;
	LRMAXDEC : LREAL;
	LRMAXVEL : LREAL;
	LRTARGETACC : LREAL;
	LRTARGETVEL : LREAL;
	LRTARGETPOS : LREAL;
	LRJERKACC : LREAL;
	LRJERKDEC : LREAL;
	LRJERKTIMEACC : LREAL;
	LRJERKTIMEDEC : LREAL;
	T5 : LREAL;
	T7 : LREAL;
END_VAR
VAR_IN_OUT
	SCPROFILEDATA : L_MB1P_ProfileData;
END_VAR
END_METHOD

METHOD CALCPROFILE_80A0_A0GTAMAX_SEARCHTIMEST5T7 : BOOL
VAR_INPUT
	LRSTARTACC : LREAL;
	LRSTARTVEL : LREAL;
	LRMAXACC : LREAL;
	LRMAXDEC : LREAL;
	LRMAXVEL : LREAL;
	LRTARGETACC : LREAL;
	LRTARGETVEL : LREAL;
	LRTARGETPOS : LREAL;
	LRJERKACC : LREAL;
	LRJERKDEC : LREAL;
	LRJERKTIMEACC : LREAL;
	LRJERKTIMEDEC : LREAL;
	T5_STARTVALUE : LREAL;
	T7_STARTVALUE : LREAL;
END_VAR
VAR_OUTPUT
	T5 : LREAL;
	T7 : LREAL;
END_VAR
END_METHOD

METHOD CALCPROFILE_80A0_A0LTAMAXT5T7 : BOOL
VAR_INPUT
	LRSTARTACC : LREAL;
	LRSTARTVEL : LREAL;
	LRMAXACC : LREAL;
	LRMAXDEC : LREAL;
	LRMAXVEL : LREAL;
	LRTARGETACC : LREAL;
	LRTARGETVEL : LREAL;
	LRTARGETPOS : LREAL;
	LRJERKACC : LREAL;
	LRJERKDEC : LREAL;
	LRJERKTIMEACC : LREAL;
	LRJERKTIMEDEC : LREAL;
	T5 : LREAL;
	T7 : LREAL;
END_VAR
VAR_IN_OUT
	SCPROFILEDATA : L_MB1P_ProfileData;
END_VAR
END_METHOD

METHOD CALCPROFILE_80A0_A0LTAMAX_SEARCHTIMEST5T7 : BOOL
VAR_INPUT
	LRSTARTACC : LREAL;
	LRSTARTVEL : LREAL;
	LRMAXACC : LREAL;
	LRMAXDEC : LREAL;
	LRMAXVEL : LREAL;
	LRTARGETACC : LREAL;
	LRTARGETVEL : LREAL;
	LRTARGETPOS : LREAL;
	LRJERKACC : LREAL;
	LRJERKDEC : LREAL;
	LRJERKTIMEACC : LREAL;
	LRJERKTIMEDEC : LREAL;
	T5_STARTVALUE : LREAL;
	T7_STARTVALUE : LREAL;
END_VAR
VAR_OUTPUT
	T5 : LREAL;
	T7 : LREAL;
END_VAR
END_METHOD

METHOD CALCPROFILE_80B0 : BOOL
VAR_INPUT
	LRSTARTACC : LREAL;
	LRSTARTVEL : LREAL;
	LRMAXACC : LREAL;
	LRMAXDEC : LREAL;
	LRMAXVEL : LREAL;
	LRTARGETACC : LREAL;
	LRTARGETVEL : LREAL;
	LRTARGETPOS : LREAL;
	LRJERKACC : LREAL;
	LRJERKDEC : LREAL;
	LRJERKTIMEACC : LREAL;
	LRJERKTIMEDEC : LREAL;
	SCMAXPROFILEDATA : L_MB1P_IntProfileData;
	SCMINPROFILEDATA : L_MB1P_IntProfileData;
END_VAR
VAR_OUTPUT
	DWSTATE : DWORD;
END_VAR
VAR_IN_OUT
	SCPROFILEDATA : L_MB1P_ProfileData;
	SCPROFILEPARAMETER : L_MB1P_ProfileParameter;
END_VAR
END_METHOD

METHOD CALCPROFILE_80B0_A0GTAMAX_SEARCHTIMEST5T7 : BOOL
VAR_INPUT
	LRSTARTACC : LREAL;
	LRSTARTVEL : LREAL;
	LRMAXACC : LREAL;
	LRMAXDEC : LREAL;
	LRMAXVEL : LREAL;
	LRTARGETACC : LREAL;
	LRTARGETVEL : LREAL;
	LRTARGETPOS : LREAL;
	LRJERKACC : LREAL;
	LRJERKDEC : LREAL;
	LRJERKTIMEACC : LREAL;
	LRJERKTIMEDEC : LREAL;
	T5_STARTVALUE : LREAL;
	T7_STARTVALUE : LREAL;
END_VAR
VAR_OUTPUT
	T5 : LREAL;
	T7 : LREAL;
END_VAR
END_METHOD

METHOD CALCPROFILE_80B0_A0GTAMAXT5T7 : BOOL
VAR_INPUT
	LRSTARTACC : LREAL;
	LRSTARTVEL : LREAL;
	LRMAXACC : LREAL;
	LRMAXDEC : LREAL;
	LRMAXVEL : LREAL;
	LRTARGETACC : LREAL;
	LRTARGETVEL : LREAL;
	LRTARGETPOS : LREAL;
	LRJERKACC : LREAL;
	LRJERKDEC : LREAL;
	LRJERKTIMEACC : LREAL;
	LRJERKTIMEDEC : LREAL;
	T5 : LREAL;
	T7 : LREAL;
END_VAR
VAR_IN_OUT
	SCPROFILEDATA : L_MB1P_ProfileData;
END_VAR
END_METHOD

METHOD CALCPROFILE_80B0_A0LTAMAXT5T7 : BOOL
VAR_INPUT
	LRSTARTACC : LREAL;
	LRSTARTVEL : LREAL;
	LRMAXACC : LREAL;
	LRMAXDEC : LREAL;
	LRMAXVEL : LREAL;
	LRTARGETACC : LREAL;
	LRTARGETVEL : LREAL;
	LRTARGETPOS : LREAL;
	LRJERKACC : LREAL;
	LRJERKDEC : LREAL;
	LRJERKTIMEACC : LREAL;
	LRJERKTIMEDEC : LREAL;
	T5 : LREAL;
	T7 : LREAL;
END_VAR
VAR_IN_OUT
	SCPROFILEDATA : L_MB1P_ProfileData;
END_VAR
END_METHOD

METHOD CALCPROFILE_80B0_A0LTAMAX_SEARCHTIMEST5T7 : BOOL
VAR_INPUT
	LRSTARTACC : LREAL;
	LRSTARTVEL : LREAL;
	LRMAXACC : LREAL;
	LRMAXDEC : LREAL;
	LRMAXVEL : LREAL;
	LRTARGETACC : LREAL;
	LRTARGETVEL : LREAL;
	LRTARGETPOS : LREAL;
	LRJERKACC : LREAL;
	LRJERKDEC : LREAL;
	LRJERKTIMEACC : LREAL;
	LRJERKTIMEDEC : LREAL;
	T5_STARTVALUE : LREAL;
	T7_STARTVALUE : LREAL;
END_VAR
VAR_OUTPUT
	T5 : LREAL;
	T7 : LREAL;
END_VAR
END_METHOD

METHOD CALCPROFILE_80C0 : BOOL
VAR_INPUT
	LRSTARTACC : LREAL;
	LRSTARTVEL : LREAL;
	LRMAXACC : LREAL;
	LRMAXDEC : LREAL;
	LRMAXVEL : LREAL;
	LRTARGETACC : LREAL;
	LRTARGETVEL : LREAL;
	LRTARGETPOS : LREAL;
	LRJERKACC : LREAL;
	LRJERKDEC : LREAL;
	LRJERKTIMEACC : LREAL;
	LRJERKTIMEDEC : LREAL;
	SCMAXPROFILEDATA : L_MB1P_IntProfileData;
	SCMINPROFILEDATA : L_MB1P_IntProfileData;
END_VAR
VAR_OUTPUT
	DWSTATE : DWORD;
END_VAR
VAR_IN_OUT
	SCPROFILEDATA : L_MB1P_ProfileData;
	SCPROFILEPARAMETER : L_MB1P_ProfileParameter;
END_VAR
END_METHOD

METHOD CALCPROFILE_80C0_SEARCHTIMEST5T7 : BOOL
VAR_INPUT
	LRSTARTACC : LREAL;
	LRSTARTVEL : LREAL;
	LRMAXACC : LREAL;
	LRMAXDEC : LREAL;
	LRMAXVEL : LREAL;
	LRTARGETACC : LREAL;
	LRTARGETVEL : LREAL;
	LRTARGETPOS : LREAL;
	LRJERKACC : LREAL;
	LRJERKDEC : LREAL;
	LRJERKTIMEACC : LREAL;
	LRJERKTIMEDEC : LREAL;
	T5_STARTVALUE : LREAL;
	T7_STARTVALUE : LREAL;
END_VAR
VAR_OUTPUT
	T5 : LREAL;
	T7 : LREAL;
END_VAR
END_METHOD

METHOD CALCPROFILE_80C0_A0LTAMAXT5T7 : BOOL
VAR_INPUT
	LRSTARTACC : LREAL;
	LRSTARTVEL : LREAL;
	LRMAXACC : LREAL;
	LRMAXDEC : LREAL;
	LRMAXVEL : LREAL;
	LRTARGETACC : LREAL;
	LRTARGETVEL : LREAL;
	LRTARGETPOS : LREAL;
	LRJERKACC : LREAL;
	LRJERKDEC : LREAL;
	LRJERKTIMEACC : LREAL;
	LRJERKTIMEDEC : LREAL;
	T5 : LREAL;
	T7 : LREAL;
END_VAR
VAR_IN_OUT
	SCPROFILEDATA : L_MB1P_ProfileData;
END_VAR
END_METHOD

METHOD CALCPROFILE_80D0 : BOOL
VAR_INPUT
	LRSTARTACC : LREAL;
	LRSTARTVEL : LREAL;
	LRMAXACC : LREAL;
	LRMAXDEC : LREAL;
	LRMAXVEL : LREAL;
	LRTARGETACC : LREAL;
	LRTARGETVEL : LREAL;
	LRTARGETPOS : LREAL;
	LRJERKACC : LREAL;
	LRJERKDEC : LREAL;
	LRJERKTIMEACC : LREAL;
	LRJERKTIMEDEC : LREAL;
	SCMAXPROFILEDATA : L_MB1P_IntProfileData;
	SCMINPROFILEDATA : L_MB1P_IntProfileData;
END_VAR
VAR_OUTPUT
	DWSTATE : DWORD;
END_VAR
VAR_IN_OUT
	SCPROFILEDATA : L_MB1P_ProfileData;
	SCPROFILEPARAMETER : L_MB1P_ProfileParameter;
END_VAR
END_METHOD

METHOD CALCPROFILE_80D0_SEARCHTIMEST5T7 : BOOL
VAR_INPUT
	LRSTARTACC : LREAL;
	LRSTARTVEL : LREAL;
	LRMAXACC : LREAL;
	LRMAXDEC : LREAL;
	LRMAXVEL : LREAL;
	LRTARGETACC : LREAL;
	LRTARGETVEL : LREAL;
	LRTARGETPOS : LREAL;
	LRJERKACC : LREAL;
	LRJERKDEC : LREAL;
	LRJERKTIMEACC : LREAL;
	LRJERKTIMEDEC : LREAL;
	T5_STARTVALUE : LREAL;
	T7_STARTVALUE : LREAL;
END_VAR
VAR_OUTPUT
	T5 : LREAL;
	T7 : LREAL;
END_VAR
END_METHOD

METHOD CALCPROFILE_80D0_A0LTAMAXT5T7 : BOOL
VAR_INPUT
	LRSTARTACC : LREAL;
	LRSTARTVEL : LREAL;
	LRMAXACC : LREAL;
	LRMAXDEC : LREAL;
	LRMAXVEL : LREAL;
	LRTARGETACC : LREAL;
	LRTARGETVEL : LREAL;
	LRTARGETPOS : LREAL;
	LRJERKACC : LREAL;
	LRJERKDEC : LREAL;
	LRJERKTIMEACC : LREAL;
	LRJERKTIMEDEC : LREAL;
	T5 : LREAL;
	T7 : LREAL;
END_VAR
VAR_IN_OUT
	SCPROFILEDATA : L_MB1P_ProfileData;
END_VAR
END_METHOD

METHOD CALCPROFILE_80E0 : BOOL
VAR_INPUT
	LRSTARTACC : LREAL;
	LRSTARTVEL : LREAL;
	LRMAXACC : LREAL;
	LRMAXDEC : LREAL;
	LRMAXVEL : LREAL;
	LRTARGETACC : LREAL;
	LRTARGETVEL : LREAL;
	LRTARGETPOS : LREAL;
	LRJERKACC : LREAL;
	LRJERKDEC : LREAL;
	LRJERKTIMEACC : LREAL;
	LRJERKTIMEDEC : LREAL;
	SCMAXPROFILEDATA : L_MB1P_IntProfileData;
	SCMINPROFILEDATA : L_MB1P_IntProfileData;
END_VAR
VAR_OUTPUT
	DWSTATE : DWORD;
END_VAR
VAR_IN_OUT
	SCPROFILEDATA : L_MB1P_ProfileData;
	SCPROFILEPARAMETER : L_MB1P_ProfileParameter;
END_VAR
END_METHOD

METHOD CALCPROFILE_80E0_PROFILEDATA : BOOL
VAR_INPUT
	LRSTARTACC : LREAL;
	LRSTARTVEL : LREAL;
	LRMAXACC : LREAL;
	LRMAXDEC : LREAL;
	LRMAXVEL : LREAL;
	LRTARGETACC : LREAL;
	LRTARGETVEL : LREAL;
	LRTARGETPOS : LREAL;
	LRJERKACC : LREAL;
	LRJERKDEC : LREAL;
	LRJERKTIMEACC : LREAL;
	LRJERKTIMEDEC : LREAL;
	T5 : LREAL;
	T7 : LREAL;
END_VAR
VAR_IN_OUT
	SCPROFILEDATA : L_MB1P_ProfileData;
END_VAR
END_METHOD

METHOD CALCPROFILE_80E0_SEARCHTIMEST5T7 : BOOL
VAR_INPUT
	LRSTARTACC : LREAL;
	LRSTARTVEL : LREAL;
	LRMAXACC : LREAL;
	LRMAXDEC : LREAL;
	LRMAXVEL : LREAL;
	LRTARGETACC : LREAL;
	LRTARGETVEL : LREAL;
	LRTARGETPOS : LREAL;
	LRJERKACC : LREAL;
	LRJERKDEC : LREAL;
	LRJERKTIMEACC : LREAL;
	LRJERKTIMEDEC : LREAL;
	T5_STARTVALUE : LREAL;
	T7_STARTVALUE : LREAL;
END_VAR
VAR_OUTPUT
	T5 : LREAL;
	T7 : LREAL;
END_VAR
END_METHOD

METHOD CALCPROFILE_80F0 : BOOL
VAR_INPUT
	LRSTARTACC : LREAL;
	LRSTARTVEL : LREAL;
	LRMAXACC : LREAL;
	LRMAXDEC : LREAL;
	LRMAXVEL : LREAL;
	LRTARGETACC : LREAL;
	LRTARGETVEL : LREAL;
	LRTARGETPOS : LREAL;
	LRJERKACC : LREAL;
	LRJERKDEC : LREAL;
	LRJERKTIMEACC : LREAL;
	LRJERKTIMEDEC : LREAL;
	SCMAXPROFILEDATA : L_MB1P_IntProfileData;
	SCMINPROFILEDATA : L_MB1P_IntProfileData;
END_VAR
VAR_OUTPUT
	DWSTATE : DWORD;
END_VAR
VAR_IN_OUT
	SCPROFILEDATA : L_MB1P_ProfileData;
	SCPROFILEPARAMETER : L_MB1P_ProfileParameter;
END_VAR
END_METHOD

METHOD CALCPROFILE_80F0_PROFILEDATA : BOOL
VAR_INPUT
	LRSTARTACC : LREAL;
	LRSTARTVEL : LREAL;
	LRMAXACC : LREAL;
	LRMAXDEC : LREAL;
	LRMAXVEL : LREAL;
	LRTARGETACC : LREAL;
	LRTARGETVEL : LREAL;
	LRTARGETPOS : LREAL;
	LRJERKACC : LREAL;
	LRJERKDEC : LREAL;
	LRJERKTIMEACC : LREAL;
	LRJERKTIMEDEC : LREAL;
	T5 : LREAL;
	T7 : LREAL;
END_VAR
VAR_IN_OUT
	SCPROFILEDATA : L_MB1P_ProfileData;
END_VAR
END_METHOD

METHOD CALCPROFILE_80F0_SEARCHTIMEST5T7 : BOOL
VAR_INPUT
	LRSTARTACC : LREAL;
	LRSTARTVEL : LREAL;
	LRMAXACC : LREAL;
	LRMAXDEC : LREAL;
	LRMAXVEL : LREAL;
	LRTARGETACC : LREAL;
	LRTARGETVEL : LREAL;
	LRTARGETPOS : LREAL;
	LRJERKACC : LREAL;
	LRJERKDEC : LREAL;
	LRJERKTIMEACC : LREAL;
	LRJERKTIMEDEC : LREAL;
	T5_STARTVALUE : LREAL;
	T7_STARTVALUE : LREAL;
END_VAR
VAR_OUTPUT
	T5 : LREAL;
	T7 : LREAL;
END_VAR
END_METHOD

(* ---- L_MB1P_POSPROFILERCLUTCH.pou ---- *)
FUNCTION_BLOCK L_MB1P_POSPROFILERCLUTCH
VAR_INPUT
	XENABLE : BOOL;
	XSYNCPOS : BOOL;
	XEXECUTEGAP : BOOL;
	XAUXEXECUTEGAP : BOOL;
	LRTASKCYCLETIME : LREAL := 0.001;
	LRSLAVESYNCOUTPOS : LREAL;
	LRCYCMASTERPOS : LREAL;
	LRCYCMASTERVEL : LREAL;
	LRCYCMASTERACC : LREAL;
	LRSETSLAVEPOS : LREAL;
	LRSETSLAVEVEL : LREAL;
	LRSETSLAVEACC : LREAL;
	LRJERK : LREAL := 10000;
	LRMAXACC : LREAL := 100;
	LRMAXDEC : LREAL := 100;
	LRMAXVEL : LREAL := 10;
END_VAR
VAR_OUTPUT
	XBUSY : BOOL;
	XDONE : BOOL;
	XACCDECSYNC : BOOL;
	XPOSSYNCHRONISED : BOOL;
	XERROR : BOOL;
	EERRORID : WORD;
	LRSETSLAVEPOSOUT : LREAL;
	LRSETSLAVEVELOUT : LREAL;
	LRSETSLAVEACCOUT : LREAL;
END_VAR
VAR
	FB_POSPROFILERPOS : L_MC1P_PosProfiler;
	SCPROFILEPARAMETER : L_MC1P_ProfileParameter;
	WSTEPPER : WORD;
	XEXECUTEPOSPROFILER : BOOL;
	LRSLAVESYNCOUTPOS_INT : LREAL;
	XAUXEXECUTEPROFILE : BOOL;
	XEXECUTEPROFILE : BOOL;
	LRSETPOSPROFILER : LREAL;
	LRSETACCPROFILER : LREAL;
	LRSETVELPROFILER : LREAL;
	LRCYCMASTERPOS_INT : LREAL;
	LRCYCMASTERVEL_INT : LREAL;
	LRCYCMASTERACC_INT : LREAL;
	XPOSSYNCHRONISED_INT : BOOL;
	XEXECUTEGAPOLD : BOOL;
	XAUXEXECUTEGAPOLD : BOOL;
	XENABLEOLD : BOOL;
	LRCYCMASTERPOS_OLD : LREAL;
	LRTOLERANCE : LREAL;
END_VAR
END_FUNCTION_BLOCK

METHOD CALL_ERRORHANDLER
END_METHOD

METHOD CALL_FBMETHODES
END_METHOD

METHOD CALL_FB_POSPROFILERPOS
END_METHOD

METHOD CALL_FB_POSPROFILERPOSINPUTS
END_METHOD

METHOD CALL_OUTPUTS
END_METHOD

METHOD CALL_PROFILEPARAMETER
END_METHOD

METHOD CALL_RESETCOMMANDS
END_METHOD

METHOD CALL_RESETOUTPUTS
END_METHOD

METHOD CALL_STATEMACHINE
END_METHOD

(* ---- L_MB1P_POSPROFILERCLUTCHSTATE.pou ---- *)
FUNCTION_BLOCK L_MB1P_POSPROFILERCLUTCHSTATE EXTENDS L_MB1P_PosProfilerClutch
VAR_INPUT
	XSYNCOUTINSTANT : BOOL;
	XMOVETOTARGETPOS : BOOL;
	LRTARGETPOS : LREAL;
	EDIRECTION : L_MC2P_ClutchDirection := L_MC2P_ClutchDirection.mcCurrentDirection;
	LRAXESCYCLELENGTH : LREAL := 360;
	EAXESTRAVERSINGRANGE : L_MC1P_TraversingRange;
	LRPOSITIONINGJERK : LREAL;
	LRPOSITIONINGACC : LREAL;
	LRPOSITIONINGDEC : LREAL;
	LRPOSITIONINGVEL : LREAL;
	LRSYNCOUTINSTANTJERK : LREAL;
	LRSYNCOUTINSTANTDEC : LREAL;
	ROVERRIDEVEL : REAL := 1.0;
	ROVERRIDEACC : REAL := 1.0;
	ROVERRIDEDEC : REAL := 1.0;
END_VAR
VAR_OUTPUT
	XREVERSING : BOOL;
	XPOSITIONING : BOOL;
	XINPOSITION : BOOL;
END_VAR
VAR
	XREVERSING_INT : BOOL;
	WMODE : WORD;
	XSYNCOUTINSTANT_OLD : BOOL;
	XMOVETOTARGETPOS_OLD : BOOL;
	XPOSMODE_INT : BOOL;
	LRTASKCYCLETIME_INT : LREAL;
	LRAXESCYCLELENGTH_INT : LREAL;
	LRTARGETPOS_INT : LREAL;
	LRTARGETPOS_LOCK : LREAL;
	LRTOLERANCEVEL : LREAL;
	LRTOLERANCEACC : LREAL;
	LRACCDIST : LREAL;
	XVELTRACE : BOOL;
	WVELTRACESTEPPER : WORD;
	LRSETACC_PROFILERPOS : LREAL;
	LRPOSPROFILERSPEED_ABS : LREAL;
	WREVERSINGVELMODE : WORD;
	LRVELZERROTOLERANZ : LREAL;
	LRSETSLAVEVELOUT_OLD : LREAL;
END_VAR
END_FUNCTION_BLOCK

METHOD CALL_CALCTARGETPOS
VAR_INPUT
	LRTARGETPOS : LREAL;
END_VAR
END_METHOD

METHOD CALL_CALCTOLERANCE
END_METHOD

METHOD CALL_CALCLRCYCMASTERPOS
END_METHOD

METHOD CALL_ERRORHANDLER
END_METHOD

METHOD CALL_FBMETHODES
END_METHOD

METHOD CALL_FB_POSPROFILERPOS
END_METHOD

METHOD CALL_FB_POSPROFILERPOSINPUTS
END_METHOD

METHOD CALL_OUTPUTS
END_METHOD

METHOD CALL_PROFILEPARAMETER
END_METHOD

METHOD CALL_PROFILEPARAMETERACCDECINMODE2
END_METHOD

METHOD CALL_RESETCOMMANDS
END_METHOD

METHOD CALL_RESETOUTPUTS
END_METHOD

METHOD CALL_STATEMACHINE
END_METHOD

(* ---- L_MB1P_PREPARATIONPATH_LM.pou ---- *)
FUNCTION_BLOCK L_MB1P_PREPARATIONPATH_LM
VAR_INPUT
	XEXECUTE : BOOL;
	XSINGLESTEP : BOOL;
	ALRSTARTPOSITION : ARRAY [1..12] OF LREAL;
	LRSTARTBLENDINGRADIUS : LREAL;
	XSTARTHALT : BOOL;
	LRPATHJERK : LREAL;
	XECOCPUMODE : BOOL;
END_VAR
VAR_OUTPUT
	XERROR : BOOL;
	EERRORID : L_IE1P_Error;
	XBUSY : BOOL;
	XDONE : BOOL;
	BYNUMOFPOINTS : BYTE;
	BYNUMOFHALT : BYTE;
	AXHALT : ARRAY [0..10] OF BOOL;
	ALRPROFILEPOINTS : ARRAY [1..10] OF ARRAY [1..12] OF LREAL;
	EENDCOORDSYSTEM : L_MC4P_CoordSystem := L_MC4P_CoordSystem.MCS;
	ALRENDPOSITION : ARRAY [1..12] OF LREAL;
	LRENDBLENDINGRADIUS : LREAL;
	XENDHALT : BOOL;
END_VAR
VAR_IN_OUT
	AXESGROUP : AXES_GROUP_KIN;
	ASCPROFILEPAR : ARRAY [1..10] OF L_TT1P_scProfilePar;
	MC_MOVELINABS : ARRAY [1..10] OF MC_MoveLinearAbsolute;
END_VAR
VAR
	WSTATE : WORD := 0;
	AXCALCPATHLEGTHBETWEENPOINTS : ARRAY [1..11] OF BOOL;
	ALRPATHLEGTHBETWEENPOINTS : ARRAY [1..11] OF LREAL;
	XSINGLESTEP_INT : BOOL;
	LRBLENDINGRADIUS_INT : LREAL;
	BYNUMOFPOINTS_LOCK : BYTE;
	XCALCINTERMEDIANTEPOINT : BOOL;
	XCPUECOMODEEXECUTE : BOOL;
	IPOINTNO : INT;
	IFORCNT : INT;
	IFORCNT2 : INT;
	LRTMP : LREAL;
	LRTMP1 : LREAL;
	LRTMP2 : LREAL;
	XERRORINVALIDPROFILE : BOOL;
	XERROR_INVALIDCOORDSYSTEM : BOOL;
	XERROR_INTERNAL : BOOL;
	XEXECUTE_OLD : BOOL;
	C_BYMAXTARGETPOINTS : BYTE := 10;
END_VAR
END_FUNCTION_BLOCK

METHOD CALL_ERRORHANDLER
END_METHOD

METHOD CALL_FBMETHODS
END_METHOD

METHOD CALL_OUTPUT
END_METHOD

METHOD CALL_RESETCOMMANDS
END_METHOD

METHOD CALL_RESETFB
END_METHOD

METHOD CALL_RESETOUTPUT
END_METHOD

METHOD CALL_STATEMACHINE
END_METHOD

METHOD GET_LRTARTGETPOSITION : LREAL
VAR_INPUT
	IAXISID : INT;
	IPOINTNO : INT;
END_VAR
END_METHOD

METHOD CALL_INIT
END_METHOD

(* ---- L_MB1P_SIMPLEPOSABORTCORRECTION.pou ---- *)
FUNCTION_BLOCK L_MB1P_SIMPLEPOSABORTCORRECTION
VAR_INPUT
	XENABLE : BOOL;
	LRCYCLETIME : LREAL;
	XABORTFROMPOSCTRL : BOOL;
	LRMAXACC : LREAL;
	LRACTVELFROMPOSCTRL : LREAL;
	LRSIMPLEPOSUNLIMITED : LREAL;
END_VAR
VAR_OUTPUT
	XABORTPROFILEFINISHED : BOOL;
	LRPOSOUT : LREAL;
END_VAR
VAR
	T_NORM_FAK : LREAL;
	T_NORM : LREAL;
	T_REAL : LREAL;
	LRSTARTPOS : LREAL;
	LRSTARTVEL : LREAL;
	R_EDGE_ABORTFROMPOSCTRL : R_TRIG;
	F_EDGE_ABORTFROMPOSCTRL : F_TRIG;
END_VAR
END_FUNCTION_BLOCK

(* ---- L_MB1P_SIMPLEPOSBASE.pou ---- *)
FUNCTION_BLOCK L_MB1P_SIMPLEPOSBASE
VAR_INPUT
	XENABLE : BOOL;
	XEXECUTE : BOOL;
	XABORTPROFILE : BOOL;
	LRCORRECTION : LREAL;
	LRMAXVELPOS : LREAL := 10;
	LRMAXVELNEG : LREAL := 10;
	LRACCDEC : LREAL := 100;
	EPROFILETYPE : L_MB1P_ProfileType := 0;
END_VAR
VAR_OUTPUT
	LRPOSOUTUNLIMITED : LREAL;
	LRRESIDUALOFFSET : LREAL;
	LRSPEEDOUT : LREAL;
	XPROFILEFAILED : BOOL;
	XPROFILEABORTED : BOOL;
	XINTARGET : BOOL;
	XBUSY : BOOL;
	DISTATE : DINT;
END_VAR
VAR_IN_OUT
	AXIS : Axis_REF;
END_VAR
VAR
	L_SDINTEGRATE1 : L_USPP_Integrate;
	R_TRIG1 : R_TRIG;
	R_TRIG2 : R_TRIG;
	F_TRIG2 : F_TRIG;
	F_TRIG3 : F_TRIG;
	DWPOSMODE : DWORD := 1;
	DWDISABLEMODE : DWORD;
	LRRAMPDISTANCE : LREAL;
	LRDELTAY : LREAL;
	LRBASICPOSITION : LREAL;
	BYSTEP : BYTE;
	BNEGSPEEDSELECTED : BOOL;
	LRXNORM : LREAL;
	LRPOSOUTOLD : LREAL;
	N : INT;
	LRMAXSPEEDINTERN : LREAL;
	LRMAXSPEEDNEG : LREAL;
	LRMAXSPEEDPOS : LREAL;
	LRSTARTPOSITION : LREAL;
	XSAVESTARTPOSITION : BOOL;
	LRPOSOUT : LREAL;
	LRPOSOUTOLDTEST : LREAL;
	LRPOSTEST : LREAL;
	XENDOFPROFILE : BOOL;
END_VAR
END_FUNCTION_BLOCK

METHOD A01_PROFILECONTROL
END_METHOD

METHOD A02_POLYNOMIAL4THORDER
END_METHOD

METHOD A03_POLYNOMIAL2NDORDER
END_METHOD

METHOD A04_POLYNOMIAL5THORDER
END_METHOD

(* ---- L_MB1P_SIMPLEPOSSETOFFSET.pou ---- *)
FUNCTION_BLOCK L_MB1P_SIMPLEPOSSETOFFSET
VAR_INPUT
	XENABLE : BOOL;
	LRCYCMASTERPOS : LREAL;
	LRCYCMASTERVEL : LREAL;
	LRCYCMASTERACC : LREAL;
	LRSETOFFSET : LREAL;
	XLOADOFFSET : BOOL;
	DWNUMERATOR : DWORD := 1;
	DWDENOMINATOR : DWORD := 1;
	EDIRECTION : L_TF1P_Direction;
	EPROFILETYPE : L_MB1P_ProfileType := 0;
	LRVELPOS : LREAL := 100.0;
	LRVELNEG : LREAL := 100.0;
	LRACCDEC : LREAL := 1000.0;
END_VAR
VAR_OUTPUT
	XBUSY : BOOL;
	XDONE : BOOL;
	XERROR : BOOL;
	EERRORID : WORD;
	LROFFSET : LREAL;
	LRSETOFFSETVELOUT : LREAL;
END_VAR
VAR_IN_OUT
	MASTERAXIS : AXIS_REF;
	SLAVEAXIS : AXIS_REF;
END_VAR
VAR
	WSTATEMASHINESIMPLEPOS : WORD := 0;
	LRSMDELTAPOS : LREAL;
	LRSIMPLEPOSOFFSET : LREAL;
	LRSALVEVELBAND : LREAL;
	LRABORTSTARTVEL : LREAL;
	LRSMSETOFFSET_OLD : LREAL;
	LRFACTOR : LREAL;
	LRLOADRESTOFFSET_INT : LREAL;
	LRVELPOS_INT : LREAL := 100.0;
	LRVELNEG_INT : LREAL := 100.0;
	LRACCDEC_INT : LREAL := 1000.0;
	XERRORINVALIDVELPOS : BOOL;
	XERRORINVALIDVELNEG : BOOL;
	XERRORINVALIDACCDEC : BOOL;
	XENABLE_OLD : BOOL;
	LROFFSET_OLD : LREAL;
	SIMPLEPOSITIONING : L_MB1P_SimplePosBase;
	ABORTPOSCTRLCORRECT : L_MB1P_SimplePosAbortCorrection;
END_VAR
END_FUNCTION_BLOCK

METHOD CALL_CALCFACTOR
END_METHOD

METHOD CALL_ERRORHANDLER
END_METHOD

METHOD CALL_FBMETHODS
END_METHOD

METHOD CALL_OUTPUT
END_METHOD

METHOD CALL_RESETCOMMANDS
END_METHOD

METHOD CALL_RESETOUTPUT
END_METHOD

METHOD CALL_SIMPLEPOS
END_METHOD

METHOD CALL_SIMPLEPOS_ABORTPOSCTRLCORRECT
END_METHOD

METHOD CALL_SIMPLEPOS_OFFSET
END_METHOD

METHOD CALL_STATEMASHINE
END_METHOD

(* ---- L_MB1P_STACK.pou ---- *)
FUNCTION_BLOCK L_MB1P_STACK
VAR_INPUT
	XENABLE : BOOL;
	XLOADTPPOS : BOOL;
	XLOADCYCSETPOS : BOOL;
	XTAKEPOS : BOOL;
	LRTPPOS : LREAL;
	LRCYCSETPOS : LREAL;
	LRCYCSETVEL : LREAL;
	LRPERIOD : LREAL;
	LRMINTPDIST : LREAL;
END_VAR
VAR_OUTPUT
	XBUSY : BOOL;
	XSTACKISFULL : BOOL;
	XSTACKISEMPTY : BOOL;
	LRPOSOUT : LREAL;
	LRDISTOUT : LREAL;
	LRSETDISTOUT : LREAL;
	XPOSPERIODOVERRUNPOS : BOOL;
	XPOSPERIODOVERRUNNEG : BOOL;
	UISTACKSTARTPOS : UINT := 0;
	UISTACKFILLSTATE : UINT := 0;
	ALRSTACKSAVEPOS : ARRAY [1..gc_uiStackLength] OF LREAL;
	AUIPERIODCNTRPOS : ARRAY [1..gc_uiStackLength] OF UINT;
	UIPERIODCNTR : UINT;
	LRTPDIST : LREAL;
	XPOSRECEIVED : BOOL;
	XPOSOUTOFWINDOW : BOOL;
	XWINDOWOPEN : BOOL;
END_VAR
VAR
	XSTACKVALUEVALID : BOOL;
	LRLATESTSAVEPOS : LREAL;
	UILATESTPERIODCNTRPOS : UINT;
	UICTR : UINT := 0;
	UIVARTEMP : UINT;
	XENABLE_OLD : BOOL;
	XLOADTPPOS_OLD : BOOL;
	XLOADCYCSETPOS_OLD : BOOL;
	XTAKEPOS_OLD : BOOL;
	XFIRSTLOADPOS : BOOL;
	LRCYCSETPOS_SAVE : LREAL;
	LRSETPOSDIFF : LREAL;
	XTAKEPOS_ACTIVE : BOOL;
	LRTEMPDIST : LREAL;
	LRCYCSETPOS_OLD : LREAL;
	FB_CHECKMODULOOVERRUN : L_MB1P_CheckModuloOverrun;
	GC_UISTACKLENGTH : UINT := 100;
END_VAR
END_FUNCTION_BLOCK

METHOD CALL_CNTRMODULOOVERRUN
VAR_IN_OUT
	LRCYCSETPOS : LREAL;
END_VAR
END_METHOD

METHOD CALL_FB_CHECKMODULOOVERRUN
VAR_IN_OUT
	LRCYCSETPOS : LREAL;
	LRCYCSETVEL : LREAL;
END_VAR
END_METHOD

METHOD CALL_RESETCOMMANDS
END_METHOD

METHOD CALL_RESETOUTPUT
END_METHOD

METHOD CALL_STACK
END_METHOD

METHOD CALL_STACK_LOADPOS
VAR_IN_OUT
	LRCYCPOS : LREAL;
	LRLOADPOS : LREAL;
END_VAR
END_METHOD

METHOD CALL_STACK_TAKEPOS
VAR_IN_OUT
	LRCYCPOS : LREAL;
END_VAR
END_METHOD

METHOD FUN_PERIODCNTRDIFF : LREAL
VAR_INPUT
	UIDIFF : UINT;
END_VAR
VAR_OUTPUT
	IOUT : INT;
END_VAR
END_METHOD

METHOD GET_LRLATESTDIST : LREAL
VAR_IN_OUT
	LRCYCPOS : LREAL;
END_VAR
END_METHOD

METHOD GET_LRTAKEPOS : LREAL
VAR_IN_OUT
	LRCYCPOS : LREAL;
END_VAR
END_METHOD

METHOD REVOKETAKEPOS
END_METHOD

METHOD SET_CYCSETPOS
VAR_IN_OUT
	LRCYCPOS : LREAL;
END_VAR
END_METHOD

METHOD SET_TPPOS
VAR_IN_OUT
	LRCYCPOS : LREAL;
	LRLOADTPPOS : LREAL;
END_VAR
END_METHOD

(* ---- L_MB1P_TPAVERAGEDIFF.pou ---- *)
FUNCTION_BLOCK L_MB1P_TPAVERAGEDIFF
VAR_INPUT
	XENABLE : BOOL;
	BYNROFCYCLES : BYTE := 20;
	XTPRECEIVED : BOOL;
	LRSETTPDIFFERENCE : LREAL;
	XTPERRORLIMITED : BOOL;
	LRSETMARKDISTANCE : LREAL;
	LRSETMAXAVERAGE : LREAL := 100;
END_VAR
VAR_OUTPUT
	LRTPERRORAVERAGE : LREAL;
	XAVERAGELIMITED : BOOL;
	LROPTIMISEDGEARFACTOR : LREAL;
END_VAR
VAR
	LRPROCENT : LREAL;
	BYNROFCYCLESINTERNAL : BYTE;
	XTPRECEIVEDOLD : BOOL;
	LRTOTALERROR : LREAL;
	BYCOUNTER : BYTE;
	LROPTIMIZATIONUNCLAMPED : LREAL;
END_VAR
END_FUNCTION_BLOCK

(* ---- L_MB1P_TPCALCDIFF.pou ---- *)
FUNCTION_BLOCK L_MB1P_TPCALCDIFF
VAR_INPUT
	XENABLE : BOOL;
	XTPRECEIVED : BOOL;
	LRACTTPPOSIN : LREAL;
	LRSETTPPOSIN : LREAL;
	LRSETMARKDISTANCE : LREAL;
END_VAR
VAR_OUTPUT
	XINITDONE : BOOL;
	XTPRECEIVEDOUT : BOOL;
	LRTPDIFFERENCE : LREAL;
	LRTPDIFFTOTAL : LREAL;
END_VAR
VAR
	XTPRECEIVEDOLD : BOOL;
END_VAR
END_FUNCTION_BLOCK

(* ---- L_MB1P_TPCONVERTTP.pou ---- *)
FUNCTION_BLOCK L_MB1P_TPCONVERTTP
VAR_INPUT
	XENABLE : BOOL;
	XTPRECEIVE : BOOL;
	LRACTTPPOSIN : LREAL;
	LRDELAYACTSET : LREAL;
	LRCYCPOSTPAXIS : LREAL;
	LRCYCPOSTARGETAXIS : LREAL;
	LRCYCLELENGTHTPAXIS : LREAL;
	LRCYCLELENGTHTARGETAXIS : LREAL;
END_VAR
VAR_OUTPUT
	XTPRECEIVED : BOOL;
	LRTPACTPOS : LREAL;
	XERROR : BOOL;
	EERRORID : L_IE1P_Error;
END_VAR
VAR
	LRPOSFIFOX : ARRAY [1..20] OF LREAL := [10(0)];
	LRPOSFIFOREG : ARRAY [1..20] OF LREAL := [10(0)];
	BYCOUNTER : INT := 1;
	LRSTACKDIFFERENCE : LREAL;
	LRTPDELTAINMS : LREAL;
	LRDELTAPCT : LREAL;
	XTPRECEIVEDOLD : BOOL;
	LRPOSDIFFTPAXIS : LREAL;
	IDIRECTION : INT;
	LRACTTPPOSIN_OLD : LREAL;
	XWAIT : BOOL;
	XWAIT_OLD : BOOL;
	LRACTTPPOSIN_INT : LREAL;
	R_TRIG1 : R_TRIG;
	BYCOMPENSATIONCYCLES : BYTE;
	LRDELAYACTSETRESIDUAL : LREAL;
	LRDELTATARGETAXIS : LREAL;
END_VAR
END_FUNCTION_BLOCK

METHOD SEARCHINSTACKNEGATIVE
END_METHOD

METHOD SEARCHINSTACKPOSITIVE
END_METHOD

(* ---- L_MB1P_TPLIMITDIFF.pou ---- *)
FUNCTION_BLOCK L_MB1P_TPLIMITDIFF
VAR_INPUT
	XTPRECEIVED : BOOL;
	LRSETTPDIFFERENCE : LREAL;
	LRSETLIMITMIN : LREAL := -100;
	LRSETLIMITMAX : LREAL := 100;
	LRSETTPWINDOW : LREAL := 2;
END_VAR
VAR_OUTPUT
	XTPRECEIVEDOUT : BOOL;
	XLIMITACTIVE : BOOL;
	XTPINWINDOW : BOOL;
	LRTPDIFFERENCELIM : LREAL;
END_VAR
VAR
	XTPRECEIVEDOLD : BOOL;
	XINITDONE : BOOL;
END_VAR
END_FUNCTION_BLOCK

(* ---- L_MB1P_TPVIRTUALACTPOS.pou ---- *)
FUNCTION_BLOCK L_MB1P_TPVIRTUALACTPOS
VAR_INPUT
	XTPWINDOWOPEN : BOOL;
	XTPRECEIVEDIN : BOOL;
	XMAXTPNOTDETECTED : BOOL;
	LRSETTPPOSIN : LREAL;
	LRACTTPPOSIN : LREAL;
END_VAR
VAR_OUTPUT
	XTPRECEIVEDOUT : BOOL;
	LRACTTPPOS : LREAL;
END_VAR
VAR
	XTPRECEIVEDINOLD : BOOL;
	XFLAGWINDOWOPENANDNOTP : BOOL := FALSE;
	XWINDOWOPENOLD : BOOL;
	XVIRTUALTPACTIVE : BOOL;
END_VAR
END_FUNCTION_BLOCK

(* ---- L_MB1P_WINDERIDENTDIAMETER.pou ---- *)
FUNCTION_BLOCK L_MB1P_WINDERIDENTDIAMETER
VAR_INPUT
	XEXECUTE : BOOL;
	XABORT : BOOL;
	XDANCERMINPOS : BOOL;
	LRACTREELSPEEDIN : LREAL;
	LRACTDANCERPOSIN : LREAL;
	XLINEVELDIAMCALC : BOOL;
	LRSETLINEVELDIAMCALC : LREAL;
	LRMAXDANCERPOS : LREAL;
	LRDANCERMATERIALLENGTH : LREAL;
	LRMAXDIAM : LREAL;
	LRDIAMCALCDIST : LREAL;
	WIDENTDIAMCALCCYCLES : WORD := 1;
	LRTASKCYCLE : LREAL := 0.001;
	LRIDENTVEL : LREAL;
	LRIDENTACC : LREAL;
	LRIDENTDEC : LREAL;
	LRIDENTJERK : LREAL;
END_VAR
VAR_OUTPUT
	XERROR : BOOL;
	EERRORID : WORD;
	XBUSY : BOOL;
	XDONE : BOOL;
	XCOMMANDABORTED : BOOL;
	LRSETREELSPEEDOUT : LREAL;
	LRIDETDIAM : LREAL;
END_VAR
VAR
	WSTATE : WORD;
	LRTASKCYCLE_INT : LREAL := 0.001;
	LRMAXDIAM_INT : LREAL;
	LRREELSPEEDFAKTOR_INT : LREAL;
	LRMAXDANCERPOS_INT : LREAL;
	LRDANCERMATERIALLENGTH_INT : LREAL;
	XLINEVELDIAMCALC_INT : BOOL;
	LRREELSPEEDOUT_INT : LREAL;
	LRACTREELDIST_INT : LREAL;
	LRACTDIST_INT : LREAL;
	LRPROFGENDIST_INT : LREAL;
	LRSETDIST_INT : LREAL;
	LRSETDISTCALCDIAM_INT : LREAL;
	LRPROFGENSTARTPOSIDENTDIAM_INT : LREAL;
	LRPROFGENENDPOSIDENTDIAM_INT : LREAL;
	LRRAMPGENDECDIST : LREAL;
	XRAMPGENHALT : BOOL;
	XIDENTSTARTVALUESVALID : BOOL;
	XIDENTENDVALUESVALID : BOOL;
	LRDANCERPOSSTARTIDENT : LREAL;
	LRDANCERPOSENDIDENT : LREAL;
	LRLINEVELSTARTIDENT : LREAL;
	LRLINEVELENDIDENT : LREAL;
	LRLINEDIST : LREAL;
	LRWNDPOSSTARTIDENT : LREAL;
	LRWNDPOSENDIDENT : LREAL;
	LRIDETNWINDDIST : LREAL;
	XERROR_INVALIDMAXDIAM : BOOL;
	XERROR_INVALIDDANCERMATERIALLENGTH : BOOL;
	XERROR_ACTDANPOSBIGGERMAXDANPOS : BOOL;
	XERROR_ACTDANPOSBIGGERMAXDANPOS_TMP : BOOL;
	XEXECUTE_OLD : BOOL;
	XABORT_OLD : BOOL;
	FB_RAMPGENERATOR1 : L_MC1P_RampGenerator;
END_VAR
END_FUNCTION_BLOCK

METHOD CALL_ERRORHANDLER
END_METHOD

METHOD CALL_FBMETHODS
END_METHOD

METHOD CALL_FB_RAMPGENERATOR
END_METHOD

METHOD CALL_OUTPUT
END_METHOD

METHOD CALL_RESETCOMMANDS
END_METHOD

METHOD CALL_RESETOUTPUT
END_METHOD

METHOD CALL_STATEMACHINE
END_METHOD

(* ---- L_MB1P_WINDERSYNCHRONISELINE.pou ---- *)
FUNCTION_BLOCK L_MB1P_WINDERSYNCHRONISELINE
VAR_INPUT
	XENABLE : BOOL;
	XSYNCLINEVEL : BOOL;
	XLOADSTARTREELSPEED : BOOL;
	LRSTARTREELSPEED : LREAL;
	LRGROUNDREELSPEED : LREAL;
	LRCYCLINEVEL : LREAL := 0;
	LRSETDIAMETER : LREAL;
	LRACC : LREAL := 1000;
	LRDEC : LREAL := 1000;
	LRJERK : LREAL := 100000;
	XMATERIALFEEDING : BOOL := FALSE;
END_VAR
VAR_OUTPUT
	XERROR : BOOL;
	EERRORID : WORD;
	XBUSY : BOOL;
	XSYNCHRONISED : BOOL;
	XACCDECSYNC : BOOL;
	LRSETREELSPEEDOUT : LREAL;
END_VAR
VAR
	WSTATE : WORD;
	LRREELSPEEDOUT_INT : LREAL;
	FB_RAMPGENERATOR1 : L_MC1P_RampGenerator;
	XENABLE_OLD : BOOL;
	XMATERIALFEEDING_OLD : BOOL;
	LRSCALEFAKTOR : LREAL;
	LRSCALEFAKTORABS : LREAL;
	WPARMODE : WORD;
	XTMP : BOOL;
END_VAR
END_FUNCTION_BLOCK

METHOD CALL_ERRORHANDLER
END_METHOD

METHOD CALL_FBMETHODS
END_METHOD

METHOD CALL_FB_RAMPGENERATOR
END_METHOD

METHOD CALL_OUTPUT
END_METHOD

METHOD CALL_RESETCOMMANDS
END_METHOD

METHOD CALL_RESETOUTPUT
END_METHOD

METHOD CALL_SETPARMODE
END_METHOD

METHOD CALL_STATEMACHINE
END_METHOD

(* ---- L_T01S_PHASECORRECTIONVEL.pou ---- *)
FUNCTION_BLOCK L_T01S_PHASECORRECTIONVEL
VAR_INPUT
	XENABLE : BOOL;
	XEXECUTECORRECTION : BOOL;
	LRCYCSETVEL : LREAL;
	LRSETCORRECTION : LREAL;
	LRCORRECTIONDISTANCE : LREAL;
END_VAR
VAR_OUTPUT
	XBUSY : BOOL;
	XCORRECTIONBUSY : BOOL;
	LRSETVELOUT : LREAL;
	LRSETCORRVELOUT : LREAL;
	LRSETPOSCORROUT : LREAL;
	XERROR : BOOL;
	EERRORID : L_IE1P_Error;
END_VAR
VAR
	LRDELTAPOSTOTAL : LREAL;
	LRMASTERDISTANCE : LREAL;
	LRPOSITIONSET : LREAL;
	LRPOSITIONNORMED : LREAL;
	LRPOSITIONOUTNORMED : LREAL;
	LRDELTAPOSCORRECTION : LREAL;
	LRPOSITIONSETOLD : LREAL;
	BYSTEPPER : BYTE;
	LRCORRECTIONDISTANCELOCAL : LREAL;
	LRCORRECTIONLOCAL : LREAL;
	LRDELTAPOSOUT : LREAL;
	XEXECUTECORRECTIONINTERN : BOOL;
	LRTASKCYCLE : LREAL;
	XINIT : BOOL := TRUE;
	INTEGRATE1 : L_USPP_Integrate;
END_VAR
END_FUNCTION_BLOCK

(* ---- L_TF1P_ADDPROFILEPICKANDPLACE.pou ---- *)
FUNCTION_BLOCK L_TF1P_ADDPROFILEPICKANDPLACE
VAR_INPUT
	XENABLE : BOOL;
	XEXECUTEPICKANDPLACE : BOOL;
	XADDPROFILE : BOOL;
	XRESETTARGETSTACK : BOOL;
	XACKPATHHALT : BOOL;
	XABORT : BOOL;
	XNOTCOORDINATEDSTOPALL : BOOL;
	XSINGLESTEP : BOOL;
	LRGRIPPERTIME : LREAL;
	LRPATHJERK : LREAL;
	LRNUMTASKCYCLESBEFOREEXECUTENEXTPROFILE : LREAL := 50;
	XCALCPROFILEMOVEPATH : BOOL;
END_VAR
VAR_OUTPUT
	XERROR : BOOL;
	XWARNING : BOOL;
	EERRORID : L_IE1P_Error;
	XBUSY : BOOL;
	XACTIVE : BOOL;
	XDONE : BOOL;
	XCOMMANDABORTED : BOOL;
	XENDOFPROFILE : BOOL;
	XTARGETSTACKISFULL : BOOL;
	XPATHHOLD : BOOL;
	XPROFILEINPREPARATION : BOOL;
	ISETPROFILENOOUT : INT;
	IPROFILEPOINTPASSED : INT;
	ITARGETPROFILEPOINT : INT;
	ALRTARGETPOSITION : ARRAY [1..12] OF LREAL;
	ESETSEGMENTTYPEOUT : L_MC4P_SegmentType;
	BYNUMOFPOINTSINPROFILE : BYTE;
	BYNUMOFHALTINPROFILE : BYTE;
	LRPATHPREPARATIONTIME : LREAL;
	LRPRECALCPROFILETIME : LREAL;
	XPROFILERESTTIMEVALID : BOOL;
	LRPROFILERESTTIME : LREAL;
	LRINTERRUPTPATHACC : LREAL;
	XLASTACTIVESEGMENT : BOOL;
	XNOACTIVESEGMENT : BOOL;
	XGRIPPERCTRLACTIVE : BOOL;
	XPULSEGRIPPER : BOOL;
	XPATHINTERRUPTOUT : BOOL;
	PAFB_MOVELINABS : POINTER TO ARRAY [1..10] OF L_MC4P_MoveLinearAbsolute_Internal;
	IMOVEPPNO : INT;
	IMOVELINNO : INT;
	PAFB_MOVELINABS1 : POINTER TO ARRAY [1..10] OF L_MC4P_MoveLinearAbsolute_Internal;
	PAFB_MOVELINABS2 : POINTER TO ARRAY [1..10] OF L_MC4P_MoveLinearAbsolute_Internal;
	PAFB_MOVELINABS3 : POINTER TO ARRAY [1..10] OF L_MC4P_MoveLinearAbsolute_Internal;
	XWAITDISABLEMOVECONTPATH : BOOL;
END_VAR
VAR_IN_OUT
	FB_EXTERNALMEMORY : L_MC4P_PickAndPlaceMemory;
	AXESGROUP : AXES_GROUP_KIN;
	ASCPROFILEPAR : ARRAY [1..10] OF L_TT1P_scProfilePar;
END_VAR
VAR
	LWTCHECKSUM_INT : LWORD;
	WSTATE : WORD;
	XSTATEMASHINEBUSY : BOOL;
	XSTATEMASHINEWAIT : BOOL;
	XSTATEMASHINEPATHHOLD : BOOL;
	XMOVEPAPSTATUSSEPPERENTRY : BOOL;
	WMOVEPAPSTATUSSEPPER_OLD : WORD;
	WMOVEPAPSTATUSSEPPER : WORD;
	REQUESTSINFO : DWORD;
	REQUESTSINFO_OLD : DWORD;
	DWRTRIG : DWORD;
	DWFTRIG : DWORD;
	EBUFFERMODEBLENDING_INT : MC_BUFFER_MODE := MC_BUFFER_MODE.mcBlendingLow;
	LRTEMP1 : LREAL;
	LRTEMP2 : LREAL;
	IDX1 : INT;
	IDX2 : INT;
	IDX3 : INT;
	UIDX1 : UINT;
	WDX1 : WORD;
	TTMP1 : TIME;
	WTMP1 : WORD;
	IFOR : INT;
	IFOREND : INT;
	ALRTARGETPOSTMP : ARRAY [1..12] OF LREAL;
	XCOUNTUPPROFILENOOUT : BOOL;
	XERRORINVALIDPROFILE : BOOL;
	XERROR_INVALIDCOORDSYSTEM : BOOL;
	XERROR_INVALIDTARGET : BOOL;
	XERROR_INVALIDPATHPAR : BOOL;
	XWARNING_TARGETSTATCKISFULL : BOOL;
	XWARNING_NOTREADYFORADDPROFILE : BOOL;
	XERROR_FB_MOVEPICKANDPLACE : BOOL;
	EERRORID_FB_MOVEPICKANDPLACE : L_IE1P_Error;
	XERROR_INTERNAL : BOOL;
	XERRORINTERNAL_INVALIDPPFBACTIVE : BOOL;
	WINTERNALERRORID_INT : WORD;
	XSINGLESTEP_LOCK : BOOL;
	LRGRIPPERTIME_LOCK : LREAL;
	XCALLFM : BOOL;
	LRTASKCYCLE : LREAL;
	LRTASKCYCLE_INV : LREAL;
	LRTIMEBEFOREEXECUTENEXTPROFILE : LREAL;
	FB_STACKTARGET : L_MC1P_StackControlArray := STRUCT(iMaxLegth := ciNumOfTargetInArray);
	ALRTARGETGRIPPERTIME : ARRAY [1..ciNumOfTargetInArray] OF LREAL;
	ALRPATHJERK : ARRAY [1..ciNumOfTargetInArray] OF LREAL;
	AXTARGETGRIPPERTIMEVALID : ARRAY [1..ciNumOfTargetInArray] OF BOOL;
	AXSINGLESTEP_INT : ARRAY [1..ciNumOfTargetInArray] OF BOOL;
	XNEWTARGET : BOOL;
	XAXESGROUPNOTREADYFORMOTION : BOOL;
	XNEXTPROFILEVALID : BOOL;
	XMOVEPPPATHINTERRUPTOUT : BOOL;
	IGRIPPERMOVEPPNO : INT;
	XPREPARENEXTPROFILE : BOOL;
	XPATHACTIVE_INT : BOOL;
	XPATHBUSY_INT : BOOL;
	XPATHDONE_INT : BOOL;
	XPATHHOLD_INT : BOOL;
	XPATHHOLDONENDHALT_INT : BOOL;
	XPATHINTERRUPTOUT_INT : BOOL;
	XPATHCOMMANDABORTED_INT : BOOL;
	XCOMMANDABORTED_INT : BOOL;
	XCOMMANDABORTE_INT : BOOL;
	XPROFILEINPREPARATION_INT : BOOL;
	LRPRECALCRESTTIMEALLSEGMENTS_INT : LREAL;
	XPRECALCPROFILERESTTIMEALLSEGMENTSVALID_INT : BOOL;
	XPRECALCPROFILERESTTIMEVALID_INT : BOOL;
	LRPRECALCPROFILERESTTIME_INT : LREAL;
	LRIPOTIME : LREAL;
	LRPATHPREPARATIONTIME_INT : LREAL;
	INUMOFACTIVEPATHSEGMENT_INT : INT;
	ICNTRACKPATHHALT_INT : INT;
	XVALIDSTARTPOS : BOOL;
	XSTARTPOINTINHALT_INT : BOOL;
	ALRSTARTPOS_INT : ARRAY [1..12] OF LREAL;
	ESTARTCOORDSYSTEM_INT : L_MC4P_CoordSystem;
	LRSTARTBLENDINGRADIUS_INT : LREAL;
	XSAVEPROFILE_INT : BOOL;
	ISAVEPROFILEEXECUTED_INT : INT;
	ISAVEPROFILESTACKSTARTPOS_INT : INT;
	ISAVEPROFILESTACKLEGTH_INT : INT;
	FB_STACKMOVEPICKANDPALCE : L_MC1P_StackControlArray := STRUCT(iMaxLegth := ciNumOfFBMovePickAndPlace);
	AIPROFILENOSTATIC : ARRAY [1..ciNumOfFBMovePickAndPlace] OF INT;
	FB_MOVEPICKANDPLACE : ARRAY [1..ciNumOfFBMovePickAndPlace] OF L_MB1P_MovePickAndPlaceState;
	CINUMOFTARGETINARRAY : INT := 10;
	CINUMOFTARGETINARRAYSETWARNING : INT := 8;
	CINUMOFFBMOVEPICKANDPLACE : INT := 3;
	EBUFFERMODEBLENDING : MC_BUFFER_MODE;
	LWTCHECKSUM : LWORD;
END_VAR
END_FUNCTION_BLOCK

METHOD CALL_ALLOCPOINTADR
END_METHOD

METHOD CALL_CALCPROFILETIME
END_METHOD

METHOD CALL_DISABLEMOVECONTPATH
VAR_IN_OUT
	AXESGROUP : AXES_GROUP_KIN;
END_VAR
END_METHOD

METHOD CALL_ERRORHANDLER
END_METHOD

METHOD CALL_FBMETHODS
END_METHOD

METHOD CALL_FB_MOVEPICKANDPLACE
END_METHOD

METHOD CALL_FB_MOVEPICKANDPLACE_STATUS
END_METHOD

METHOD CALL_GRIPPERCONTROL
END_METHOD

METHOD CALL_OUTPUT
END_METHOD

METHOD CALL_REQUESTS_EXT
END_METHOD

METHOD CALL_RESETCOMMANDS
END_METHOD

METHOD CALL_RESETOUTPUT
END_METHOD

METHOD CALL_STATEMACHINE
END_METHOD

METHOD CALL_ABORTPROFILE
END_METHOD

METHOD CALL_READSTARTPOSITION
END_METHOD

METHOD CALL_SAVEPROFILE
END_METHOD

METHOD CALL_TARGETSTAICPOSSTACK
END_METHOD

METHOD CALL_SETPROFILE
END_METHOD

METHOD GET_ALRINTERMEDIANTEPOINT
VAR_IN_OUT
	ALRINTERMEDIANTEPOINT : ARRAY [1..12] OF LREAL;
END_VAR
END_METHOD

METHOD CALL_INIT
END_METHOD

METHOD CALL_S000_CYCLIC
END_METHOD

(* ---- L_TF1P_REGISTERCONTROLBASE.pou ---- *)
FUNCTION_BLOCK L_TF1P_REGISTERCONTROLBASE
VAR_INPUT
	XENABLE : BOOL;
	XSYNCPOS : BOOL;
	LRVELIN : LREAL;
	LRACTSETPOSSLAVE : LREAL;
	XMARKRECEIVE : BOOL;
	ETPMODE : L_TF1P_TpMode;
	LRCYCPOSEXTENCODER : LREAL;
	LRCYCLELENGTHEXTENCODER : LREAL;
	LRACTMARKPOSIN : LREAL;
	XLOADREGPOS : BOOL;
	LRLOADREGPOS : LREAL;
	LRMARKSENSORPOS : LREAL;
	LRMARKDIST : LREAL;
	LRMAXCORRNEG : LREAL;
	LRMAXCORRPOS : LREAL;
	ESOURCEFORCORRWINDOW : L_TT1P_SourceForCorrWindow;
	LRUPPERCORRPOS : LREAL;
	LRLOWERCORRPOS : LREAL;
	DNNUMAXISY : DWORD;
	DNDENAXISY : DWORD;
	XSYNCHRONISED : BOOL;
	LRTPAXISCOMPFACTOR : LREAL;
	LRTPAXISDELAYCYCLE : LREAL;
END_VAR
VAR_OUTPUT
	LRPOSOUT : LREAL;
	LRACTVEL : LREAL;
	XERROR : BOOL;
	WERRORID : WORD;
	XLIMITACTIVE : BOOL;
	LRACTMARKERROR : LREAL;
	LRACTMARKDIST : LREAL;
	XINITDONE : BOOL;
	XCORRACTIVE : BOOL;
	XMARKRECEIVED : BOOL;
	LRREGMARKPOS : LREAL;
	XCORRNEXTCYCLE : BOOL;
END_VAR
VAR_IN_OUT
	MASTERAXIS : AXIS_REF;
	SLAVEAXIS : AXIS_REF;
END_VAR
VAR
	SPEEDTOPOSINTEGRATE : L_MC1P_IntegrateAxis;
	TPLIMITDIFF : L_MB1P_TpLimitDiff;
	FB_ADDOFFSET : L_MC1P_AddOffsetCyclic;
	TPCALCDIFF : L_MC1P_TpCalcDiff;
	CONVERTTPPOSITION : L_TT1P_CalculateTPOnMaterialPos := STRUCT(xNoMarkStack := TRUE);
	DISTCORRECTIONWINDOW : L_MB1P_DistCorrectionWindow;
	LRGEARINGFAKTOR : LREAL := 1.0;
	XERROR_TM : BOOL;
	EERRORID_TM : L_IE1P_Error;
	LRTPDIFFERENCE_INT : LREAL;
	XLOADMARKSENSORPOS_OLD : BOOL;
	XTPRECEIVED_OLD : BOOL;
	LRMARKWINDOWSIZE_INT : LREAL;
	XTPINWINDOW : BOOL;
	LRPOS_INT : LREAL;
	XTPRECEIVEDOUT_INT : BOOL;
	LRTPACTPOSITION_INT : LREAL;
	LRTPDIFFERENCELIM_INT : LREAL;
	LROFFSETPOSCTRL_INT : LREAL;
	LRPOSOUT_INT : LREAL;
	LRVELOUT_INT : LREAL;
	XCORRACTIVE_INT : BOOL;
	XINIT : BOOL := TRUE;
	XTPCORRECTIONACTIVE : BOOL := FALSE;
	LRTPAXISSETPOS : LREAL;
	LRMARKDIST_INT : LREAL;
	XZERO : BOOL;
	XHOMINGDONE : BOOL;
	XSTARTREFERENCEACTIVE : BOOL;
	XHOMINGACTIVE : BOOL := FALSE;
	XMARKDISTCHANGED : BOOL;
	XENABLE_OLD : BOOL;
	XTPRECEIVEDOUT_INTOLD : BOOL;
	XSTARTFIRSTCORRECTION : BOOL;
	LRTPDIFFERENCELIM2_INT : LREAL;
	XCORRECTIONBUSYOLD : BOOL;
	LRTPACTPOSIN_OLD : LREAL;
	LRTPSETPOSIN_OLD : LREAL;
	LRCYCLELENGTH : LREAL;
	ICOUNTER : INT := 0;
	LRSETPOSITIONOLD : LREAL;
	LRCYCLELENGTHTP : LREAL;
	LRTPACTPOSITIONOLD : LREAL;
	L_MB1P_CHECKMODULOOVERRUNSETPOS : L_MB1P_CheckModuloOverrun;
	L_MB1P_CHECKMODULOOVERRUNACTPOS : L_MB1P_CheckModuloOverrun;
	BYCYCLECOUNT_INT : BYTE;
	BYCYCLECOUNTREG_INT : BYTE;
	BYSTATE : BYTE;
	ABYCYCLECOUNT : ARRAY [0..5] OF BYTE;
	BYCYCLECOUNTSUM : BYTE;
	XFIRSTTOUCHPROBE : BOOL := TRUE;
	XCORRBASEDONMASTERPOS_INT : BOOL := FALSE;
	XTPCALCDIFFTPRECEIVEDOLD : BOOL;
	LRTPDIFFERENCECOMP_INT : LREAL;
	LRTPAXISACTPOS : LREAL;
	LRTPAXISACTVELOCITY : LREAL;
	LRTPAXISCYCLELENGTH : LREAL;
	LRCYCREGISTERPOSINT : LREAL;
	LRTPACTPOSITION_ORIGINAL : LREAL;
	LRREGISTERTOUCHPROBEDIFFERENCE : LREAL;
	LRAXISTOUCHPROBEDIFFERENCE : LREAL;
END_VAR
END_FUNCTION_BLOCK

METHOD CALL_CALCACTMARKDIST
END_METHOD

METHOD CALL_CORRECTIONPOS
END_METHOD

METHOD CALL_ENABLEREGISTERCONTROL
END_METHOD

METHOD CALL_ERRORHANDLER
END_METHOD

METHOD CALL_FB
END_METHOD

METHOD CALL_GEARING
END_METHOD

METHOD CALL_INPUT
END_METHOD

METHOD CALL_LIMIT
END_METHOD

METHOD CALL_MARKDISTCHANGE
END_METHOD

METHOD CALL_NOTENABLE
END_METHOD

METHOD CALL_OUTPUT
END_METHOD

METHOD CALL_RESET
END_METHOD

METHOD CALL_TOUCHPROBE
END_METHOD

METHOD CALL_TOUCHPROBESOURCE
END_METHOD

METHOD GET_ACTUALMARKDIST : LREAL
END_METHOD

METHOD GET_CORRREGPOS : LREAL
END_METHOD

METHOD GET_INTEGRATORREGPOS : LREAL
END_METHOD

METHOD GET_MARKERRORUNLIMITED : LREAL
END_METHOD

METHOD GET_MARKPOSITIONINREGISTER : LREAL
END_METHOD

METHOD GET_MARKRECEIVEUNLIMITED : BOOL
END_METHOD

METHOD GET_REGISTERINPUTVEL : LREAL
END_METHOD

METHOD GET_SETVELOCITYREGISTER : LREAL
END_METHOD

METHOD SET_CORRECTIONONMASTERPOS
VAR_INPUT
	XCORRBASEDONMASTER : BOOL;
END_VAR
END_METHOD

(* ---- L_TF1P_REGISTERCONTROLSTATE.pou ---- *)
FUNCTION_BLOCK L_TF1P_REGISTERCONTROLSTATE EXTENDS L_TF1P_RegisterControlBase
VAR_INPUT
	LRACTOFFSETMASTERIN : LREAL;
	LRACTOFFSETSLAVEIN : LREAL;
	XTEACHMARKWINDOW : BOOL;
	LRMARKWINDOWSIZE : LREAL;
	LRSETOFFSETMARKWINDOW : LREAL;
	DWMAXNUMBERVIRTUALMARKS : DWORD;
	LRGEARFACTORCORRGAIN : LREAL;
	LRMAXGEARFACTORCORR : LREAL;
	LRSENSORTOOLDISTANCE : LREAL;
	XGEARFACTORCORR : BOOL;
	XGEARFACTORCORRHOLD : BOOL;
	XENABLETOOLCORRECTION : BOOL;
END_VAR
VAR_OUTPUT
	XMARKWINDOWOPEN : BOOL;
	XMARKOUTOFWINDOW : BOOL;
	XMARKNOTDETECTED : BOOL;
	XMARKWINDOWTEACHED : BOOL;
	LRAVERAGEGEARFACTORCORR : LREAL;
	XGEARFACTORCORRLIMITED : BOOL;
END_VAR
VAR
	MARKWINDOW : L_MB1P_MarkWindowRelative;
	MARKSTACK : L_MB1P_MarkStack;
	TPVIRTUALACTPOS : L_MB1P_TpVirtualActPos;
	LRMARKSTACKLENGTH : LREAL;
	LRTPDIFFERENCELIMITOUT_INT : LREAL;
	XTPRECEIVESTACKOUT_INT : BOOL;
	XTPNOTDETECTED_INT : BOOL;
	XMAXTPNOTDETECTED : BOOL;
	LRGEARFACTORINTEGRATOR : LREAL;
	LRGEARFACTORGAIN : LREAL := 1;
	LRGEARFACTORNUMERATORCORR : LREAL;
	LRGEARFACTORNUMERATORCORRLIMITED : LREAL;
	LRGEARFACTORDENOMINATOR : LREAL;
	LRGEARFACTORNUMERATOR : LREAL;
	LCORRECTIONVELIN : LREAL;
	LRDELTAGEARFACTORCORR : LREAL;
	XTPSENSORTEACHEDOLD : BOOL;
	XTPSENSORTEACHEDATLASTMARK : BOOL;
	XCALCMARKDISTINITIALISED : BOOL;
	XTEACHTPSENSOROLD : BOOL;
	LRTPDEADTIMEDIFF : LREAL;
	XTPRECEIVEDOUTOLD_INT : BOOL;
	XMARKSTACKTPRECEIVEDOUTOLD : BOOL;
	LRTPACTPOSITIONREGISTER_INT : LREAL;
	XTPRECEIVEDOUTREGISTER_INT : BOOL;
	XTPRECEIVEDOUTCALCERROR_INT : BOOL;
	LRTPACTPOSMARKWINDOWIN_INT : LREAL;
	LRMASTERACTPOSITIONOLD_INT : LREAL;
END_VAR
END_FUNCTION_BLOCK

METHOD CALL_AVERAGETPDIFF
END_METHOD

METHOD CALL_CALCACTMARKDIST
END_METHOD

METHOD CALL_CORRECTIONPOS
END_METHOD

METHOD CALL_ENABLEREGISTERCONTROL
END_METHOD

METHOD CALL_ERRORHANDLER
END_METHOD

METHOD CALL_FB
END_METHOD

METHOD CALL_INPUT
END_METHOD

METHOD CALL_LIMIT
END_METHOD

METHOD CALL_MARKDISTCHANGE
END_METHOD

METHOD CALL_MARKREGISTER
END_METHOD

METHOD CALL_MARKWINDOW
END_METHOD

METHOD CALL_NOTENABLE
END_METHOD

METHOD CALL_OUTPUT
END_METHOD

METHOD CALL_RESET
END_METHOD

METHOD CALL_TOUCHPROBE
END_METHOD

METHOD CALL_TOUCHPROBESOURCE
END_METHOD

METHOD CALL_VIRTUALACTPOS
END_METHOD

METHOD GET_ACTMARKERRORLIMITED : LREAL
END_METHOD

METHOD GET_MARKRECEIVEDLIMITED : BOOL
END_METHOD

METHOD GET_MARKWINDOWCOMP : BOOL
END_METHOD

METHOD GET_LRMARKSTACKLENGTH : LREAL
END_METHOD

(* ---- L_TF1P_SYNCDRIVEPOSBASE.pou ---- *)
FUNCTION_BLOCK L_TF1P_SYNCDRIVEPOSBASE
VAR_INPUT
	XENABLE : BOOL;
	LRCYCMASTERPOS : LREAL;
	LRCYCMASTERVEL : LREAL;
	LRCYCMASTERACC : LREAL;
	XLOADSTARTSLAVEPOS : BOOL := FALSE;
	LRSTARTSLAVEPOS : LREAL;
	XLOADGEARBOXPOS : BOOL;
	LRLOADGEARBOXPOS : LREAL;
	DWNUMERATOR : DWORD := 1;
	DWDENOMINATOR : DWORD := 1;
	LRSETOFFSET : LREAL;
END_VAR
VAR_OUTPUT
	XERROR : BOOL;
	EERRORID : L_IE1P_Error;
	XBUSY : BOOL;
	LRSETSLAVEPOSOUT : LREAL;
	LRSETSLAVEVELOUT : LREAL;
	LRSETSLAVEACCOUT : LREAL;
	LRSETGEARBOXPOSOUT : LREAL;
	LROFFSET : LREAL;
END_VAR
VAR_IN_OUT
	MASTERAXIS : AXIS_REF;
	SLAVEAXIS : AXIS_REF;
END_VAR
VAR
	LRSCALING_INT : LREAL := 1;
	LRGEARBOXSTARTPOSOUT_INT : LREAL;
	LRSETMASTERVEL_INT : LREAL;
	LRSETMASTERVEL_OLD : LREAL;
	LRSETMASTERACC_INT : LREAL;
	DWDENOMINATOR_INT : DWORD := 1;
	XENABLE_OLD : BOOL;
	WAXESMODE : WORD;
	ESTATE : L_TF1P_States := L_TF1P_States.INIT;
	ESTATE_OLD : L_TF1P_States := L_TF1P_States.INIT;
	XSTATEENTRY : BOOL;
	XENABLEGEARBOX : BOOL;
	FB_ADDOFFSETCYCLIC : L_MC1P_AddOffsetCyclic;
	FB_GEARBOXPOSITION : L_MB1P_GearboxPosition;
	FB_AXISCONVERTER : L_MC2P.L_MC2P_AxisConverterBase;
	LRLOADGEARBOXPOS_INT : LREAL;
	LRSETGEARBOXPOSOUT_INT : LREAL;
	LRSETGEARBOXPOSOUT_OLD : LREAL;
END_VAR
END_FUNCTION_BLOCK

METHOD CALL_AXESMODE
END_METHOD

METHOD CALL_ERRORHANDLER
END_METHOD

METHOD CALL_FBMETHODS
END_METHOD

METHOD CALL_FBMETHODS_FMDISABLE
END_METHOD

METHOD CALL_FB_ADDOFFSETCYCLIC
END_METHOD

METHOD CALL_FB_ADDOFFSETCYCLIC_INPUT
END_METHOD

METHOD CALL_FB_AXISCONVERTER
END_METHOD

METHOD CALL_FB_AXISCONVERTER_INPUT
END_METHOD

METHOD CALL_FB_GEARBOXPOSITION
END_METHOD

METHOD CALL_FB_GEARBOXPOSITION_INPUT
END_METHOD

METHOD CALL_FB_GEARBOXPOSITION_LOADGEARBOXPOS
END_METHOD

METHOD CALL_LOADSLAVESTARTPOS
END_METHOD

METHOD CALL_OUTPUT
END_METHOD

METHOD CALL_OUTPUT_OFFSET
END_METHOD

METHOD CALL_OUTPUT_SETSLAVEOUT
END_METHOD

METHOD CALL_RESETCOMMANDS
END_METHOD

METHOD CALL_RESETFM
END_METHOD

METHOD CALL_RESETOUTPUT
END_METHOD

METHOD CALL_STATEMASHINE
END_METHOD

METHOD CALL_S000_CYCLIC
END_METHOD

METHOD CALL_S001_INIT
END_METHOD

METHOD CALL_S010_READY
END_METHOD

METHOD CALL_S200_SYNCHRON
END_METHOD

METHOD CALL_S998_ERROR
END_METHOD
